      def clipWhenLowerLimitIsLessThanHigher(outputScaledValue, outputRange):
          if (outputScaledValue < outputRange[0]):
              return outputRange[0]
          elif (outputScaledValue > outputRange[1]):
              return outputRange[1]
          else:
              return outputScaledValue
          end
      end

      slope = computeSlope(rawRange, scaledRange)
      intercept = computeIntercept(slope, rawRange, scaledRange)
      scaledValue = slope * value + intercept
      return clipScaledValue(scaledValue, scaledRange)
  end

  def limit(value, range):
      return scale(value, range, range)
  end


  rq_init_comm_if_connected(9, "1")
  rq_init_comm_if_connected(2, "2")
  rq_init_comm_if_connected(3, "3")
  rq_init_comm_if_connected(4, "4")
  rq_print_connected_grippers()
  rq_gripper_communication_thread = run rq_gripper_communication()
  set_closed_norm(97.6470588235294, 1)
  set_open_norm(1.1764705882352942, 1)
  set_closed_mm(0.0, 1)
  set_open_mm(53.0, 1)
  set_closed_norm(100.0, 2)
  set_open_norm(0.0, 2)
  set_closed_mm(0.0, 2)
  set_open_mm(50.0, 2)
  set_closed_norm(100.0, 3)
  set_open_norm(0.0, 3)
  set_closed_mm(0.0, 3)
  set_open_mm(50.0, 3)
  set_closed_norm(100.0, 4)
  set_open_norm(0.0, 4)
  set_closed_mm(0.0, 4)
  set_open_mm(50.0, 4)
  rq_current_limit_enabled = False
  while(not rq_gripper_communication_thread_started):
      sync()
  end
  # end: URCap Installation Node
  # begin: URCap Installation Node
  #   Source: OPC UA, 2.0.2, Rocketfarm AS
  #   Type: OPC UA
  global opcua_daemon = rpc_factory("xmlrpc", "http://127.0.0.1:40409/RPC2")
  def opcua_client_connect(address):
  return opcua_daemon.client_connect(address)
  end
  def opcua_client_get_id(client_name):
  return opcua_daemon.client_get_id(client_name)
  end
  def opcua_client_try_connect(client_id):
  opcua_result = False
  if (opcua_daemon.client_connect(client_id)):
  sleep(0.01)
  opcua_result = opcua_daemon.client_is_connected(client_id)
  opcua_retry = 10
  while ( (not opcua_result) and (opcua_retry > 0) ):
  sleep(0.1)
  opcua_result = opcua_daemon.client_is_connected(client_id)
  opcua_retry = opcua_retry - 1
  end
  end
  return opcua_result
  end
  def opcua_client_disconnect(client_id):
  return opcua_daemon.client_disconnect(client_id)
  end
  def opcua_client_is_connected(client_id):
  return opcua_daemon.client_is_connected(client_id)
  end
  def opcua_client_read_byid(client_id, namespace_id, variable_id):
  return opcua_daemon.client_read_variable_by_id(client_id, namespace_id, variable_id)
  end
  def opcua_client_read_byname(client_id, namespace_id, variable_name):
  return opcua_daemon.client_read_variable_by_name(client_id, namespace_id, variable_name)
  end
  def opcua_client_write_byid(client_id, namespace_id, variable_id, variable_value):
  return opcua_daemon.client_write_variable_by_id(client_id, namespace_id, variable_id, variable_value)
  end
  def opcua_client_write_byname(client_id, namespace_id, variable_name, variable_value):
  return opcua_daemon.client_write_variable_by_name(client_id, namespace_id, variable_name, variable_value)
  end
  def opcua_client_last_error(client_id):
  return opcua_daemon.client_get_last_error(client_id)
  end
  def opcua_server_read_byname(variable_name):
  return opcua_daemon.server_read_variable_by_name(variable_name)
  end
  def opcua_server_write_byname(variable_name, variable_value):
  return opcua_daemon.server_write_variable_by_name(variable_name, variable_value)
  end
  def opcua_server_last_error():
  return opcua_daemon.server_get_last_error()
  end
  def opcua_error_to_string(errorCode):
  return opcua_daemon.error_code_to_string(errorCode)
  end
  # end: URCap Installation Node
  global AMR_Position=struct(position_identifier=0, x1=0, x2=0, y1=0, y2=0, theta1=0, theta2=0)
  global CAM_Pose=p[0,0,0,0,0,0]
  global CAM_Relation=""
  global CMD_Abort=  False
  global CMD_Clear=  False
  global CMD_Reset=  False
  global CMD_Start=  False
  global CMD_Suspend=  False
  global CMD_Unhold=  False
  global CMD_Unsuspend=  False
  global CNT_Rack_Output=0
  global FNC_Freedrive=  False
  global PRC_TubCounter=0
  global STP=0
  global easyPickCount=0
  global easyPickCount_4=0
  global easyPickCount_6=0
  global easyPickNoObj=0
  global easyPickNoObj_4=0
  global easyPickNoObj_6=0
  global easyPickParts=0
  global easyPickParts_4=0
  global easyPickParts_6=0
  global Container_mid_1_p=p[-.379239199143, -.127191311915, .299999999998, .000000000046, -.000000000021, -1.247199999994]
  global Container_mid_1_q=[-2.477408934449926, -1.2969853503591224, -1.875639182904262, -1.539621866126728, 1.5731943360401213, -2.8009955944022717]
  global Container_capt_p=p[-.525590029047, .407247642794, .411588185841, -.000000000107, .000000000065, -2.896148821900]
  global Container_capt_q=[-3.5968351615224767, -2.0050156108707204, -0.8176271154495112, -1.8895759482008394, 1.5730967555598792, -2.2743681102957645]
  global Waypoint_51_p=p[-.335468094724, -.217855817953, .299999999998, .000000000047, -.000000000014, -.994837065669]
  global Waypoint_51_q=[-2.2250460001249586, -1.2969853503591224, -1.875639182904262, -1.539621866126728, 1.573194336040121, -2.800995594402271]
  global Waypoint_65_p=p[-.380578560601, .136229906820, .300065486591, .002668209125, -.001950299791, -1.918285884015]
  global Waypoint_65_q=[-3.1484482924090784, -1.309784547691681, -1.8656262159347534, -1.5396564540318032, 1.5732260942459106, -2.8009706179248255]
  global Waypoint_86_p=p[-.610891912545, .328076512140, .154928874949, -.144389774448, 2.158207980619, -2.101916875088]
  global Waypoint_86_q=[-3.0298424402820032, -2.1616608105101527, -1.770405888557434, -1.8800016842284144, -0.04927570024599248, -0.4936583677874964]
  global Waypoint_16_p=p[-.530358413935, .418971000515, -.109643658887, -.463059997969, 2.087871459122, -2.058033430549]
  global Waypoint_16_q=[-3.2300904432879847, -2.6409207783141078, -1.877760410308838, -1.6937691173949183, -0.43063193956484014, 0.029483795166015625]
  global Waypoint_87_p=p[-.459488806274, .188986755628, .171097942578, -.348072585494, -2.059579317749, 2.019661285019]
  global Waypoint_87_q=[-2.790591303502218, -2.152559896508688, -1.6884642839431763, -2.469414850274557, 0.6884214878082275, 0.021232735365629196]
  global Waypoint_89_p=p[-.261886355761, -.111669623901, .131097242659, -1.173634433322, -1.227274747052, 1.193766216763]
  global Waypoint_89_q=[-2.672995464666928, -2.175407175402028, -1.7617490112425536, -2.338843663300132, 2.030865036219133, 0.036428578240585985]
  global Waypoint_90_p=p[-.269165142951, -.108082457315, .026677271969, -1.173634433324, -1.227274747052, 1.193766216762]
  global Waypoint_90_q=[-2.6853380119023815, -2.380020912479904, -1.7522585114443245, -2.1436252765786143, 2.018787725064888, 0.03659425986402358]
  global Waypoint_88_p=p[-.617446503519, .392270291627, .170489198955, -.224010410006, -2.066036920971, 2.088909130040]
  global Waypoint_88_q=[-3.1488035953258766, -2.4221038789008897, -1.1666724558911366, -2.618578428321003, 0.2380794033913185, -0.04528854192806264]
  global Waypoint_94_p=p[-.452978066378, .173533334300, .109390198136, -.002578830757, -2.196586508502, 2.177068753404]
  global Waypoint_94_q=[-2.6674557574892073, -2.1212895090252317, -1.967198705482553, -2.208419381150989, 0.5117897724834828, 0.04481344519449531]
  global Waypoint_93_p=p[-.596468537907, .142788156334, .105779109453, -.673355127215, 1.831389627653, -1.853156743314]
  global Waypoint_93_q=[-2.6921545586066635, -2.073966887503291, -2.065600898968258, -2.154852607781155, -0.22224352987151796, 0.042304121657345886]
  global Waypoint_95_p=p[-.605386387448, -.069660570533, .218481828695, .000812734400, .006677866481, -1.958478278110]
  global Waypoint_95_q=[-2.8029143834677903, -1.8400819882842256, -1.544169955118452, -1.327224466208456, 1.5676652012497132, -2.4155226342256775]
  global Waypoint_13_p=p[-.479450777041, .284140798427, .125270103493, -.276792173670, 2.098433187455, -2.121256516887]
  global Waypoint_13_q=[-2.8915050665484827, -1.9549266300597132, -2.2318272590637207, -1.6654960117735804, 0.020810842514038086, -0.4019392172442835]
  global Waypoint_70_p=p[-.472820924464, .292439826304, .207418370234, -.259787347864, -2.053484648504, 2.070709755662]
  global Waypoint_70_q=[-2.969927421603815, -2.07168115810532, -1.6835546062719366, -2.4953958198513964, 0.4489790927922641, -0.005578998612037367]
  global Waypoint_2_p=p[-.312961047461, -.152991312519, .223609826854, -.745314530454, -1.713873240489, 1.673341715282]
  global Waypoint_2_q=[-2.3560472170459192, -2.183784624139303, -1.4583134651184082, -2.6435262165465296, 1.6522362232208252, 0.043451953679323196]
  global Waypoint_3_p=p[-.113749865836, -.390110151572, .317307487562, -.519383711706, -.839884211339, 1.756868173041]
  global Waypoint_3_q=[-1.8909733931170862, -1.720626016656393, -1.5115610361099243, -2.1240560017027796, 2.1809096336364746, 0.7227501273155212]
  global Waypoint_15_p=p[.029144035010, -.436802470887, .327885032028, -.521560953301, -.623641814548, 1.862659450154]
  global Waypoint_15_q=[-1.564817253743307, -1.556895188321807, -1.6826975345611572, -1.6944714985289515, 2.2362685203552246, 1.117417335510254]
  global Waypoint_14_p=p[.068712235638, -.569419545175, .285215357659, -.679242949116, -.712065334485, 1.394044574094]
  global Waypoint_14_q=[-1.5731792953485346, -1.8029235103747094, -1.6781008808776736, -1.2218450646111982, 2.4719572998240125, 1.6394218026856375]
  global Waypoint_4_p=p[-.047220457210, -.557624911767, .136370962514, -.679242949107, -.712065334475, 1.394044574096]
  global Waypoint_4_q=[-1.7740079055958748, -2.0023561428872334, -1.7577251142892676, -1.18903287716154, 2.4487287370345143, 1.322902469273079]
  global Waypoint_25_p=p[.065436479647, -.569388431626, .287820755049, -.679242949185, -.712065334557, 1.394044574070]
  global Waypoint_25_q=[-1.5789263550890595, -1.8020194754825436, -1.6702557537748035, -1.237882536889547, 2.471995808083492, 1.6301087487321393]
  global Waypoint_39_p=p[.137772150180, -.577759956854, .299999999946, .000000000217, -.000000000207, -1.594351842625]
  global Waypoint_39_q=[-1.108978697428574, -1.776486680444405, -1.413737665315093, -1.5218908901738937, 1.5733062372356947, -1.0863866394180182]
  global Waypoint_41_p=p[.074222967010, -.565641640647, .234620140366, -.516884386806, .529223682286, -1.529619060506]
  global Waypoint_41_q=[-0.9596722604286052, -1.8767069964135548, -1.4892746174057256, -1.7813862040292285, 1.0520698599867686, -0.8199687448260349]
  global Waypoint_40_p=p[.039987741677, -.564832865048, .191055405868, -.767560686167, .343136533060, -2.241315728308]
  global Waypoint_40_q=[-1.0070649180116558, -1.8745927522477324, -1.6139175023195245, -1.6337474788493545, 1.032708081143138, -0.11587278312988403]
  global Waypoint_42_p=p[.041363380882, -.564865360786, .192805844739, .278500165520, .624117100927, .762272396553]
  global Waypoint_42_q=[-1.0050718976263102, -1.8744386685524779, -1.609151451954446, -1.6399653140247947, 1.0334006002355505, -3.254032861659603]
  global Waypoint_43_p=p[.041363380886, -.564865360780, .192805844755, .854271020883, .226833028600, 2.453002871494]
  global Waypoint_43_q=[-1.0050567614299233, -1.874341297657562, -1.6092945416026048, -1.6397580431809713, 1.0333661149462194, -5.0371728933995605]
  global Waypoint_44_p=p[.040882892233, -.564854254876, .192193763716, .110913882012, .659173708659, .275719738520]
  global Waypoint_44_q=[-1.0057704811530535, -1.8745207681598055, -1.6107765025572558, -1.637858394640876, 1.033164860873599, -2.7487836132940755]
  global Waypoint_45_p=p[.042647731639, -.564895808997, .194439423694, -.451694728506, .563172064821, -1.343350300184]
  global Waypoint_45_q=[-1.0032860829914387, -1.8741561795270565, -1.6048483308761785, -1.6453689714776623, 1.0342050634514657, -1.06078829880322]
  global Waypoint_46_p=p[.099944144487, -.566244126804, .267342790130, -.451694834765, .563172023386, -1.343350532536]
  global Waypoint_46_q=[-0.9257438092434924, -1.889970530402497, -1.3828165217629076, -1.8916791100652528, 1.0664350961373816, -0.9805910833329659]
  global Waypoint_47_p=p[.099944144444, -.566244126727, .267342790273, -.101742139519, .058679218003, -1.457888523314]
  global Waypoint_47_q=[-1.1112623176383014, -1.729989471869196, -1.5530029871033957, -1.4442770617454777, 1.4670579052775654, -1.2224020460061675]
  global Waypoint_48_p=p[-.136182767566, -.647487115908, .294247768372, -.101742139549, .058679218020, -1.457888523312]
  global Waypoint_48_q=[-1.532196177857717, -1.9115932455375173, -1.2651848069729779, -1.5055651746702665, 1.4703193777418382, -1.646379689188814]
  global Waypoint_49_p=p[-.159024328559, -.641021381179, .047691706070, -.000000000033, -.000000000027, -1.457897102937]
  global Waypoint_49_q=[-1.6098490079965062, -2.1164987141784586, -1.6156631902166785, -0.9800092198841526, 1.573231151532669, -1.722204302767242]
  global Waypoint_50_p=p[-.159024328558, -.641021381151, .291114489351, -.000000000033, -.000000000027, -1.457897102937]
  global Waypoint_50_q=[-1.609190265995684, -1.9426985888940234, -1.2189094859258596, -1.55056435122874, 1.5734384912955113, -1.7235116759964022]
  def Sub_Vision_V18():
    $ 650 "Sub_Vision_V18" "noBreak"
    $ 651 "PreSettings"
    $ 652 "CAM_LM_Detected≔ False "
    global CAM_LM_Detected=  False
    $ 653 "CAM_Captures≔0"
    global CAM_Captures=0
    $ 654 "CAM_Pose≔p[0,0,0,0,0,0]"
    global CAM_Pose=p[0,0,0,0,0,0]
    $ 655 "CAM_LM_Refinmnt≔ False "
    global CAM_LM_Refinmnt=  False
    $ 656 "CAM_LM_Refined≔ False "
    global CAM_LM_Refined=  False
    $ 657 "CAM_LM_Deviatn≔p[0,0,0,0,0,0]"
    global CAM_LM_Deviatn=p[0,0,0,0,0,0]
    $ 658 "CAM_LM_ID≔0"
    global CAM_LM_ID=0
    $ 659 "CAM_Done≔ False "
    global CAM_Done=  False
    $ 660 "CAM_CNT_Obj≔0"
    global CAM_CNT_Obj=0
    $ 661 "CAM_Result = []"
    CAM_Result = []
    $ 662 "OBJ_Detected≔ False "
    global OBJ_Detected=  False
    $ 663 "FRM_Reference≔p[0,0,0,0,0,0]"
    global FRM_Reference=p[0,0,0,0,0,0]
    $ 664 "'=========='"
    # '=========='
    $ 665 "Switch Action"
    switch_1 = Action
    $ 666 "Case 13"
    if (13 == switch_1):
    elif (15 == switch_1):
      $ 784 "Case 15"
    elif (131 == switch_1):
      $ 830 "Case 131"
      $ 831 "Read (SensoPart)"
      $ 832 "Action_Info≔'search for landmark'"
      global Action_Info="search for landmark"
      $ 833 "CAM_LM≔CAM_LMs[4]"
      global CAM_LM=CAM_LMs[4]
      $ 834 "CAM_Relation≔CAM_LM.capture_relation"
      global CAM_Relation=CAM_LM.capture_relation
      $ 835 "go to capture pose"
      $ 838 "If ITM_ID≟1 and JIG≟7"
      if (ITM_ID == 1  and  JIG == 7):
        $ 839 "PSE_T≔uLM_Cap_SSRack"
        global PSE_T=uLM_Cap_SSRack
      else:
        $ 840 "ElseIf ITM_ID≟5 and JIG≟7"
        if (ITM_ID == 5  and  JIG == 7):
          $ 841 "PSE_T≔FRM_Cap_SSRack"
          global PSE_T=FRM_Cap_SSRack
        else:
          $ 842 "ElseIf ITM_ID≟13 and JIG≟7"
          if (ITM_ID == 13  and  JIG == 7):
            $ 843 "PSE_T≔FRM_pick_rack_const"
            global PSE_T=p[-0.5568395192387274,0.34423986364170267,0.44698620470146266,-1.0069110132199915E-6,3.378712467497258E-5,-8.002029546773325E-6]
          else:
            $ 844 "ElseIf ITM_ID≟1 and JIG≟15"
            if (ITM_ID == 1 and JIG == 15):
              $ 845 "MoveJ"
              $ 846 "Container_mid_1" "breakAfter"
              movej(get_inverse_kin(Container_mid_1_p, qnear=Container_mid_1_q), a=1.3962634015954636, v=1.0471975511965976, r=0.05)
              $ 847 "Container_capt" "breakAfter"
              movej(get_inverse_kin(Container_capt_p, qnear=Container_capt_q), a=1.3962634015954636, v=1.0471975511965976)
              $ 848 "PSE_T≔FRM_Container_S_const"
              global PSE_T=p[-0.510412665574981,0.40064363362973565,0.41159789496794374,-1.1370875604168537E-5,-3.643547521609506E-6,-2.896122366208473]
            else:
              $ 849 "ElseIf ITM_ID≟1 and JIG≟16"
              if (ITM_ID == 1  and  JIG == 16):
                $ 850 "MoveJ"
                $ 851 "Waypoint_51" "breakAfter"
                movej(get_inverse_kin(Waypoint_51_p, qnear=Waypoint_51_q), a=1.3962634015954636, v=1.0471975511965976, r=0.05)
                $ 854 "PSE_T≔FRM_Container_S_const"
                global PSE_T=p[-0.510412665574981,0.40064363362973565,0.41159789496794374,-1.1370875604168537E-5,-3.643547521609506E-6,-2.896122366208473]
              else:
                $ 855 "ElseIf ITM_ID≟1 and JIG≟17"
                if (ITM_ID == 1  and  JIG == 17):
                  $ 856 "MoveJ"
                  $ 857 "Waypoint_51" "breakAfter"
                  movej(get_inverse_kin(Waypoint_51_p, qnear=Waypoint_51_q), a=1.3962634015954636, v=1.0471975511965976, r=0.05)
                  $ 860 "PSE_T≔FRM_Container_S_const"
                  global PSE_T=p[-0.510412665574981,0.40064363362973565,0.41159789496794374,-1.1370875604168537E-5,-3.643547521609506E-6,-2.896122366208473]
                else:
                  $ 861 "ElseIf ITM_ID≟1 and JIG≟18"
                  if (ITM_ID == 1  and  JIG == 18):
                    $ 864 "MoveJ"
                    $ 865 "Waypoint_51" "breakAfter"
                    movej(get_inverse_kin(Waypoint_51_p, qnear=Waypoint_51_q), a=1.3962634015954636, v=1.0471975511965976, r=0.05)
                    $ 866 "Waypoint_65" "breakAfter"
                    movej(get_inverse_kin(Waypoint_65_p, qnear=Waypoint_65_q), a=1.3962634015954636, v=1.0471975511965976)
                    $ 867 "PSE_T≔FRM_Container_S_const"
                    global PSE_T=p[-0.510412665574981,0.40064363362973565,0.41159789496794374,-1.1370875604168537E-5,-3.643547521609506E-6,-2.896122366208473]
                  else:
                    $ 868 "ElseIf ITM_ID≟1 and JIG≟19"
                    if (ITM_ID == 1  and  JIG == 19):
                      $ 871 "MoveJ"
                      $ 872 "Waypoint_51" "breakAfter"
                      movej(get_inverse_kin(Waypoint_51_p, qnear=Waypoint_51_q), a=1.3962634015954636, v=1.0471975511965976, r=0.05)
                      $ 874 "PSE_T≔aq_rack1_const"
                      global PSE_T=p[-0.6171199234912242,0.18274496130308399,0.4990241423073791,7.867082192074154E-6,-3.513408957609815E-5,-2.5093516385827686]
                    end
                  end
                end
              end
            end
          end
        end
      end
      $ 875 "do_transition(PSE_T, keep_rxry=False)"
      do_transition(PSE_T, keep_rxry=False)
      $ 876 "Set"
      set_tcp(p[0.0,0.0,0.161,3.1415,0.0,0.0])
      $ 877 "MoveJ"
      $ 878 "PSE_T" "breakAfter"
      movej(PSE_T, a=1.3962634015954636, v=1.7453292519943295)
      $ 879 "CAM_Pose≔get_actual_tcp_pose()"
      global CAM_Pose= get_actual_tcp_pose ()
      $ 880 "Loop  not CAM_Done and  not ERROR.FLAG and  not CMD_Stop"
      while (  not  CAM_Done  and    not  ERROR.FLAG  and    not  CMD_Stop):
        $ 881 "adjust capture pose"
        $ 882 "If CAM_LM_Detected and CAM_LM_Refinmnt"
        if (CAM_LM_Detected  and  CAM_LM_Refinmnt):
          $ 883 "PSE_T≔p[0,0,0.300,0,0,0]"
          global PSE_T=p[0,0,0.300,0,0,0]
          $ 884 "CAM_Pose≔PSE_T"
          global CAM_Pose=PSE_T
          $ 885 "If  not is_reachable(FRM_Reference,[PSE_T])"
          if (  not  is_reachable(FRM_Reference,[PSE_T])):
            $ 886 "Error"
            $ 887 "set_error(ERROR_POSE_NOT_REACHABLE)"
            set_error(ERROR_POSE_NOT_REACHABLE)
          end
          $ 888 "If  not ERROR.FLAG"
          if (  not  ERROR.FLAG):
            $ 889 "MoveJ"
            $ 890 "PSE_T" "breakAfter"
            set_tcp(p[0.0,0.0,0.161,0.0,0.0,0.0])
            movej(pose_trans(FRM_Reference, PSE_T), a=0.8726646259971648, v=1.3962634015954636)
            $ 891 "CAM_LM_Refined≔ True "
            global CAM_LM_Refined=  True
          end
        else:
          $ 892 "ElseIf  not CAM_LM_Detected and CAM_Captures>0"
          if (  not  CAM_LM_Detected  and  CAM_Captures>0):
            $ 893 "MoveL"
            $ 894 "If FRM_Reference≟p[0,0,0,0,0,0]"
            if (FRM_Reference == p[0,0,0,0,0,0]):
              $ 895 "PSE_T≔get_random_pose(pose_ref=CAM_Pose, mode='cubic', range_max=[0.150,0.150,0.015])"
              global PSE_T=get_random_pose(pose_ref=CAM_Pose, mode="cubic", range_max=[0.150,0.150,0.015])
            else:
              $ 900 "Else" "noBreak"
              $ 901 "PSE_T≔get_random_pose(pose_ref=CAM_Pose, mode='rotation', range_max=[10,10,0])"
              global PSE_T=get_random_pose(pose_ref=CAM_Pose, mode="rotation", range_max=[10,10,0])
              $ 902 "CAM_LM_Refined≔ True "
              global CAM_LM_Refined=  True
            end
            $ 903 "If get_inverse_kin_has_solution(pose_trans(FRM_Reference, PSE_T))"
            if (get_inverse_kin_has_solution( pose_trans (FRM_Reference, PSE_T))):
              $ 904 "Comment"
              # Comment
              $ 905 "PSE_T" "breakAfter"
              set_tcp(p[0.0,0.0,0.161,3.1415,0.0,0.0])
              movel(pose_trans(FRM_Reference, PSE_T), a=0.03, v=0.05)
            else:
              $ 906 "Else" "noBreak"
              $ 907 "'If random pose is out of reach, set the initial cam pose'"
              # 'If random pose is out of reach, set the initial cam pose'
              $ 908 "PSE_T≔CAM_Pose"
              global PSE_T=CAM_Pose
            end
          end
        end
        $ 909 "Wait: 2.0"
        sleep(2.0)
        $ 910 "trigger"
        $ 911 "If ITM_ID≟1 and JIG≟7"
        if (ITM_ID == 1  and  JIG == 7):
          # begin: URCap Program Node
          #   Source: SensoPart VISOR Robotic, 2.0.0, SensoPart Industriesensorik GmbH
          #   Type: VISOR Trigger
          $ 912 "# 1 VISOR Trigger"
          visor_changeJob(1, "Landmark_INVITE_2", 6000)
          visor_trigger(1, 6000, "arm")
          # end: URCap Program Node
        else:
          $ 913 "ElseIf ITM_ID≟5 and JIG≟7"
          if (ITM_ID == 5  and  JIG == 7):
            # begin: URCap Program Node
            #   Source: SensoPart VISOR Robotic, 2.0.0, SensoPart Industriesensorik GmbH
            #   Type: VISOR Trigger
            $ 914 "# 1 VISOR Trigger"
            visor_changeJob(1, "Landmark_INVITE_2", 6000)
            visor_trigger(1, 6000, "arm")
            # end: URCap Program Node
          else:
            $ 915 "ElseIf ITM_ID≟13 and JIG≟7"
            if (ITM_ID == 13  and  JIG == 7):
              # begin: URCap Program Node
              #   Source: SensoPart VISOR Robotic, 2.0.0, SensoPart Industriesensorik GmbH
              #   Type: VISOR Trigger
              $ 916 "# 1 VISOR Trigger"
              visor_changeJob(1, "Landmark_INVITE_2", 6000)
              visor_trigger(1, 6000, "arm")
              # end: URCap Program Node
            else:
              $ 917 "ElseIf ITM_ID≟1 and JIG≟15"
              if (ITM_ID == 1 and JIG == 15):
                # begin: URCap Program Node
                #   Source: SensoPart VISOR Robotic, 2.0.0, SensoPart Industriesensorik GmbH
                #   Type: VISOR Trigger
                $ 918 "# 1 VISOR Trigger"
                visor_changeJob(1, "PowderA", 6000)
                visor_trigger(1, 6000, "arm")
                # end: URCap Program Node
              else:
                $ 919 "ElseIf ITM_ID≟1 and JIG≟16"
                if (ITM_ID == 1 and JIG == 16):
                  # begin: URCap Program Node
                  #   Source: SensoPart VISOR Robotic, 2.0.0, SensoPart Industriesensorik GmbH
                  #   Type: VISOR Trigger
                  $ 920 "# 1 VISOR Trigger"
                  visor_changeJob(1, "Weigh_target", 6000)
                  visor_trigger(1, 6000, "arm")
                  # end: URCap Program Node
                else:
                  $ 921 "ElseIf ITM_ID≟1 and JIG≟17"
                  if (ITM_ID == 1 and JIG == 17):
                    # begin: URCap Program Node
                    #   Source: SensoPart VISOR Robotic, 2.0.0, SensoPart Industriesensorik GmbH
                    #   Type: VISOR Trigger
                    $ 922 "# 1 VISOR Trigger"
                    visor_changeJob(1, "Weigh_dispense", 6000)
                    visor_trigger(1, 6000, "arm")
                    # end: URCap Program Node
                  else:
                    $ 923 "ElseIf ITM_ID≟1 and JIG≟18"
                    if (ITM_ID == 1 and JIG == 18):
                      # begin: URCap Program Node
                      #   Source: SensoPart VISOR Robotic, 2.0.0, SensoPart Industriesensorik GmbH
                      #   Type: VISOR Trigger
                      $ 924 "# 1 VISOR Trigger"
                      visor_changeJob(1, "pick_rack", 6000)
                      visor_trigger(1, 6000, "arm")
                      # end: URCap Program Node
                    else:
                      $ 926 "ElseIf ITM_ID≟1 and JIG≟19"
                      if (ITM_ID == 1 and JIG == 19):
                        # begin: URCap Program Node
                        #   Source: SensoPart VISOR Robotic, 2.0.0, SensoPart Industriesensorik GmbH
                        #   Type: VISOR Trigger
                        $ 927 "# 1 VISOR Trigger"
                        visor_changeJob(1, "place_rack", 6000)
                        visor_trigger(1, 6000, "arm")
                        # end: URCap Program Node
                      end
                    end
                  end
                end
              end
            end
          end
        end
        $ 932 "TM_3D≔visor_partsFound(1)"
        global TM_3D= visor_partsFound (1)
        $ 933 "If TM_3D>0"
        if (TM_3D>0):
          $ 934 "CAM_LM_Detected≔ True "
          global CAM_LM_Detected=  True
          $ 935 "CAM_Captures≔0"
          global CAM_Captures=0
        else:
          $ 936 "Else" "noBreak"
          $ 937 "CAM_LM_Detected≔ False "
          global CAM_LM_Detected=  False
          $ 938 "CAM_Captures≔CAM_Captures+1"
          global CAM_Captures=CAM_Captures+1
        end
        $ 943 "result"
        $ 944 "If CAM_LM_Detected"
        if (CAM_LM_Detected):
          $ 945 "If (CAM_LM_Refinmnt and CAM_LM_Refined) or  not CAM_LM_Refinmnt"
          if ((CAM_LM_Refinmnt  and  CAM_LM_Refined)  or    not  CAM_LM_Refinmnt):
            $ 1003 "If ITM_ID≟1 and JIG≟7"
            if (ITM_ID == 1  and  JIG == 7):
              $ 1004 "CAM_LM_SSRack≔visor_getPose3d(1, 0)"
              global CAM_LM_SSRack= visor_getPose3d (1, 0)
            else:
              $ 1005 "ElseIf ITM_ID≟5 and JIG≟7"
              if (ITM_ID == 5  and  JIG == 7):
                $ 1006 "CAM_LM_SSRack≔visor_getPose3d(1, 0)"
                global CAM_LM_SSRack= visor_getPose3d (1, 0)
              else:
                $ 1007 "ElseIf ITM_ID≟13 and JIG≟7"
                if (ITM_ID == 13  and  JIG == 7):
                  $ 1008 "CAM_LM_Bott≔visor_getPose3d(1, 0)"
                  global CAM_LM_Bott= visor_getPose3d (1, 0)
                else:
                  $ 1009 "ElseIf ITM_ID≟1 and JIG≟15"
                  if (ITM_ID == 1 and JIG == 15):
                    $ 1010 "CAM_LM_Cont_S≔visor_getPose3d(1, 0)"
                    global CAM_LM_Cont_S= visor_getPose3d (1, 0)
                    $ 1011 "cont_img_pose≔get_actual_tcp_pose()"
                    global cont_img_pose= get_actual_tcp_pose ()
                  else:
                    $ 1012 "ElseIf ITM_ID≟1 and JIG≟16"
                    if (ITM_ID == 1 and JIG == 16):
                      $ 1013 "CAM_cont≔visor_getPose3d(1, 0)"
                      global CAM_cont= visor_getPose3d (1, 0)
                      $ 1014 "cont_img_pose≔get_actual_tcp_pose()"
                      global cont_img_pose= get_actual_tcp_pose ()
                    else:
                      $ 1015 "ElseIf ITM_ID≟1 and JIG≟17"
                      if (ITM_ID == 1 and JIG == 17):
                        $ 1016 "pose_rack_aq1≔visor_getPose3d(1, 0)"
                        global pose_rack_aq1= visor_getPose3d (1, 0)
                        $ 1017 "cont_img_pose≔get_actual_tcp_pose()"
                        global cont_img_pose= get_actual_tcp_pose ()
                      else:
                        $ 1018 "ElseIf ITM_ID≟1 and JIG≟18"
                        if (ITM_ID == 1 and JIG == 18):
                          $ 1019 "pose_rack_aq1≔visor_getPose3d(1, 0)"
                          global pose_rack_aq1= visor_getPose3d (1, 0)
                          $ 1020 "FRM_Container_S≔get_actual_tcp_pose()"
                          global FRM_Container_S= get_actual_tcp_pose ()
                        else:
                          $ 1021 "ElseIf ITM_ID≟1 and JIG≟19"
                          if (ITM_ID == 1 and JIG == 19):
                            $ 1022 "pose_rack_aq1≔visor_getPose3d(1, 0)"
                            global pose_rack_aq1= visor_getPose3d (1, 0)
                            $ 1023 "aq_rack1≔get_actual_tcp_pose()"
                            global aq_rack1= get_actual_tcp_pose ()
                          end
                        end
                      end
                    end
                  end
                end
              end
            end
            $ 1024 "CAM_Done≔ True "
            global CAM_Done=  True
          end
        else:
          $ 1025 "ElseIf  not CAM_LM_Detected and CAM_Captures<CAM_PRM_Retries"
          if (  not  CAM_LM_Detected  and  CAM_Captures<CAM_PRM_Retries):
            $ 1026 "CAM_LM_Refined≔ False "
            global CAM_LM_Refined=  False
          else:
            $ 1027 "ElseIf CAM_Captures≥CAM_PRM_Retries"
            if (CAM_Captures >= CAM_PRM_Retries):
              $ 1028 "CAM_Done≔ True "
              global CAM_Done=  True
              $ 1029 "Error"
              $ 1030 "set_error(ERROR_NO_LANDMARK)"
              set_error(ERROR_NO_LANDMARK)
            end
          end
        end
      end
    elif (151 == switch_1):
      $ 1031 "Case 151"
      $ 1032 "Detect (SensoPart)"
      $ 1033 "go to capture pose"
      $ 1034 "FRM_Reference≔FRM_Cap_SSRack"
      global FRM_Reference=FRM_Cap_SSRack
      $ 1035 "PSE_T≔p[0,0,-0.00,0,0,0]"
      global PSE_T=p[0,0,-0.00,0,0,0]
      $ 1036 "do_transition(pose_trans(FRM_Reference, PSE_T), keep_rxry=False)"
      do_transition( pose_trans (FRM_Reference, PSE_T), keep_rxry=False)
      $ 1037 "JNT_Q≔get_actual_joint_positions()"
      global JNT_Q= get_actual_joint_positions ()
      $ 1038 "JNT_Q≔[JNT_Q[0], JNT_Q[1], JNT_Q[2], JNT_Q[3], JNT_Q[4], 0]"
      global JNT_Q=[JNT_Q[0], JNT_Q[1], JNT_Q[2], JNT_Q[3], JNT_Q[4], 0]
      $ 1039 "Set"
      set_tcp(p[0.0,0.0,0.161,3.1415,0.0,0.0])
      $ 1040 "movej(get_inverse_kin(pose_trans(FRM_Reference, PSE_T), qnear=JNT_Q))"
      movej(get_inverse_kin( pose_trans (FRM_Reference, PSE_T), qnear=JNT_Q))
      $ 1041 "CAM_Pose≔pose_trans(pose_inv(FRM_Reference), get_actual_tcp_pose())"
      global CAM_Pose= pose_trans ( pose_inv (FRM_Reference),  get_actual_tcp_pose ())
      $ 1042 "Loop  not CAM_Done and  not ERROR.FLAG and  not CMD_Stop"
      while (  not  CAM_Done  and    not  ERROR.FLAG  and    not  CMD_Stop):
        $ 1043 "If  not OBJ_Detected and CAM_Captures>0"
        if (  not  OBJ_Detected  and  CAM_Captures>0):
          $ 1044 "MoveL"
          $ 1045 "If FRM_Reference≟p[0,0,0,0,0,0]"
          if (FRM_Reference == p[0,0,0,0,0,0]):
            $ 1047 "PSE_T≔get_random_pose(pose_ref=CAM_Pose, mode='rotation', range_max=[15,15,0])"
            global PSE_T=get_random_pose(pose_ref=CAM_Pose, mode="rotation", range_max=[15,15,0])
          else:
            $ 1048 "Else" "noBreak"
            $ 1049 "PSE_T≔get_random_pose(pose_ref=CAM_Pose, mode='rotation', range_max=[10,10,0])"
            global PSE_T=get_random_pose(pose_ref=CAM_Pose, mode="rotation", range_max=[10,10,0])
          end
          $ 1050 "If get_inverse_kin_has_solution(pose_trans(FRM_Reference, PSE_T))"
          if (get_inverse_kin_has_solution( pose_trans (FRM_Reference, PSE_T))):
            $ 1051 "PSE_T" "breakAfter"
            set_tcp(p[0.0,0.0,0.161,3.1415,0.0,0.0])
            movel(pose_trans(FRM_Reference, PSE_T), a=0.03, v=0.05)
          else:
            $ 1052 "Else" "noBreak"
            $ 1053 "'If random pose is out of reach, set the initial cam pose'"
            # 'If random pose is out of reach, set the initial cam pose'
            $ 1054 "PSE_T≔CAM_Pose"
            global PSE_T=CAM_Pose
            $ 1055 "PSE_T" "breakAfter"
            set_tcp(p[0.0,0.0,0.161,3.1415,0.0,0.0])
            movel(pose_trans(FRM_Reference, PSE_T), a=0.03, v=0.05)
          end
        end
        $ 1056 "Wait: 0.5"
        sleep(0.5)
        $ 1057 "Set"
        set_tcp(p[0.0,0.0,0.161,3.1415,0.0,0.0])
        # begin: URCap Program Node
        #   Source: SensoPart VISOR Robotic, 2.0.0, SensoPart Industriesensorik GmbH
        #   Type: VISOR Trigger
        $ 1058 "# 1 VISOR Trigger"
        visor_changeJob(1, "Object Detection Single", 6000)
        visor_trigger(1, 6000, "arm")
        # end: URCap Program Node
        $ 1059 "If visor_isResponseOk(1)"
        if ( visor_isResponseOk (1)):
          $ 1060 "CAM_CNT_Obj≔visor_partsFound(1)"
          global CAM_CNT_Obj= visor_partsFound (1)
          $ 1061 "CAM_OBJ_Pose≔visor_getPose3d(1, 0)"
          global CAM_OBJ_Pose= visor_getPose3d (1, 0)
          $ 1062 "If CAM_CNT_Obj>0"
          if (CAM_CNT_Obj>0):
            $ 1063 "CAM_OBJ_Color≔visor_getAdditionalData(1, 0)"
            global CAM_OBJ_Color= visor_getAdditionalData (1, 0)
            $ 1064 "CAM_DetectScore≔to_num(visor_getAdditionalData(1, 1))/1000"
            global CAM_DetectScore=to_num( visor_getAdditionalData (1, 1))/1000
            $ 1065 "OBJ_Detected≔ True "
            global OBJ_Detected=  True
          end
        else:
          $ 1066 "Else" "noBreak"
          $ 1067 "CAM_Captures≔CAM_Captures+1"
          global CAM_Captures=CAM_Captures+1
        end
        $ 1068 "If OBJ_Detected"
        if (OBJ_Detected):
          $ 1069 "Get object data"
          $ 1070 "PRC_CntDetect≔0"
          global PRC_CntDetect=0
          $ 1071 "Loop PRC_CntDetect<CAM_CNT_Obj"
          while (PRC_CntDetect<CAM_CNT_Obj):
            $ 1072 "get object and jig number"
            $ 1073 "If ITM_ID≟1 and JIG≟7"
            if (ITM_ID == 1  and  JIG == 7):
              $ 1074 "FRM_Reference≔FRM_Cap_SSRack"
              global FRM_Reference=FRM_Cap_SSRack
            else:
              $ 1075 "ElseIf ITM_ID≟5 and JIG≟7"
              if (ITM_ID == 5  and  JIG == 7):
                $ 1076 "FRM_Reference≔uLM_Cap_SSRack"
                global FRM_Reference=uLM_Cap_SSRack
              end
            end
            $ 1079 "PSE_T≔pose_trans(pose_inv(FRM_Reference), CAM_OBJ_Pose)"
            global PSE_T= pose_trans ( pose_inv (FRM_Reference), CAM_OBJ_Pose)
            $ 1080 "CAM_Result.append(get_pattern_counter(PSE_T, 'X', pattern=[10, 5], patternsize=[0.181, 0.081]))"
            CAM_Result.append(get_pattern_counter(PSE_T, "X", pattern=[10, 5], patternsize=[0.181, 0.081]))
            $ 1081 "PRC_CntDetect≔PRC_CntDetect+1"
            global PRC_CntDetect=PRC_CntDetect+1
          end
          $ 1082 "CAM_Done≔ True "
          global CAM_Done=  True
        else:
          $ 1083 "ElseIf CAM_Captures≥CAM_PRM_Retries"
          if (CAM_Captures >= CAM_PRM_Retries):
            $ 1084 "CAM_Done≔ True "
            global CAM_Done=  True
          else:
            $ 1085 "Else" "noBreak"
            $ 1086 "CAM_Captures≔CAM_Captures+1"
            global CAM_Captures=CAM_Captures+1
          end
        end
      end
    end
    $ 1087 "'=========='"
    # '=========='
    $ 1088 "PostSettings"
    $ 1089 "FRM_Reference≔p[0,0,0,0,0,0]"
    global FRM_Reference=p[0,0,0,0,0,0]
    $ 1090 "Set"
    set_tcp(p[0.0,0.0,0.161,3.1415,0.0,0.0])
    $ 1091 "CAM_Pose≔p[0,0,0,0,0,0]"
    global CAM_Pose=p[0,0,0,0,0,0]
    $ 1092 "Action≔0"
    global Action=0
    $ 1093 "Action_Info≔''"
    global Action_Info=""
  end
  def Sub_AMR_MiR_V3():
    $ 1094 "Sub_AMR_MiR_V3" "noBreak"
    $ 1095 "PreSettings"
    $ 1096 "AMR_TargetList≔[1,2,3,4,5,21,22,23,24,31,32,33,34,35,36,37,38,41]"
    global AMR_TargetList=[1,2,3,4,5,21,22,23,24,31,32,33,34,35,36,37,38,41]
    $ 1097 "AMR_Done≔ False "
    global AMR_Done=  False
    $ 1098 "AMR_PosActual≔T2O_Current_Pos"
    global AMR_PosActual=modbus_get_signal_status("T2O_Current_Pos")
    $ 1099 "AMR_Attemps≔T2O_Nav_Attemps"
    global AMR_Attemps=modbus_get_signal_status("T2O_Nav_Attemps")
    $ 1100 "AMR_Battery≔MiR_Battery_Lvl"
    global AMR_Battery=modbus_get_signal_status("MiR_Battery_Lvl")
    $ 1101 "AMR_Charging≔(T2O_Charging≟1)"
    global AMR_Charging=(modbus_get_signal_status("T2O_Charging") == 1)
    $ 1102 "AMR_Position≔struct(position_identifier=T2O_Current_Pos, x1=MiR_Position_X1, x2=MiR_Position_X2, y1=MiR_Position_Y1, y2=MiR_Position_Y2, theta1=MiR_Theta_1, theta2=MiR_Theta_2) "
    global AMR_Position=struct(position_identifier=modbus_get_signal_status("T2O_Current_Pos"), x1=modbus_get_signal_status("MiR_Position_X1"), x2=modbus_get_signal_status("MiR_Position_X2"), y1=modbus_get_signal_status("MiR_Position_Y1"), y2=modbus_get_signal_status("MiR_Position_Y2"), theta1=modbus_get_signal_status("MiR_Theta_1"), theta2=modbus_get_signal_status("MiR_Theta_2"))
    $ 1103 "If MiR_Mode≠7"
    if (modbus_get_signal_status("MiR_Mode") != 7):
      $ 1104 "Error"
      $ 1105 "set_error(ERROR_AMR_WRONG_MODE)"
      set_error(ERROR_AMR_WRONG_MODE)
      $ 1106 "AMR_Done≔ True "
      global AMR_Done=  True
    end
    $ 1107 "'=========='"
    # '=========='
    $ 1108 "Switch STATE"
    switch_1 = STATE
    $ 1109 "Case 1"
    if (1 == switch_1):
      $ 1110 "stopping"
      $ 1111 "If T2O_Done≟1 and O2T_Acknowledge≟0"
      if (modbus_get_signal_status("T2O_Done") == 1  and  modbus_get_signal_status("O2T_Acknowledge") == 0):
        $ 1112 "Set O2T_Acknowledge=1"
        modbus_set_output_register("O2T_Acknowledge", 1)
      end
      $ 1113 "Set MiR_CMD_Stop=On"
      modbus_set_output_signal("MiR_CMD_Stop", True)
      $ 1114 "AMR_Position.position_identifier = 0"
      AMR_Position.position_identifier = 0
      $ 1115 "AMR_Done≔ True "
      global AMR_Done=  True
    elif (2 == switch_1):
      $ 1116 "Case 2"
      $ 1117 "stopped"
      $ 1118 "If MiR_State≠3 and MiR_State≠5"
      if (modbus_get_signal_status("MiR_State") != 3  and  modbus_get_signal_status("MiR_State") != 5):
        $ 1119 "Set MiR_CMD_Stop=Off"
        modbus_set_output_signal("MiR_CMD_Stop", False)
      end
    elif (3 == switch_1):
      $ 1120 "Case 3"
      $ 1121 "resetting"
      $ 1122 "Set O2T_Mis_Main=Off"
      modbus_set_output_signal("O2T_Mis_Main", False)
      $ 1123 "Set O2T_Mis_Charge=Off"
      modbus_set_output_signal("O2T_Mis_Charge", False)
      $ 1124 "If MiR_Mis_Queue>0"
      if (modbus_get_signal_status("MiR_Mis_Queue")>0):
        $ 1125 "Set MiR_CMD_Clear_Q=On"
        modbus_set_output_signal("MiR_CMD_Clear_Q", True)
        $ 1126 "Wait MiR_Mis_Queue≟0"
        while (not(modbus_get_signal_status("MiR_Mis_Queue") == 0)):
          sync()
        end
        $ 1127 "Set MiR_CMD_Clear_Q=Off"
        modbus_set_output_signal("MiR_CMD_Clear_Q", False)
      end
      $ 1128 "If MiR_Error_ID≠0"
      if (modbus_get_signal_status("MiR_Error_ID") != 0):
        $ 1129 "Set MiR_CMD_Clear_E=On"
        modbus_set_output_signal("MiR_CMD_Clear_E", True)
        $ 1130 "Wait MiR_Error_ID≟0"
        while (not(modbus_get_signal_status("MiR_Error_ID") == 0)):
          sync()
        end
        $ 1131 "Set MiR_CMD_Clear_E=Off"
        modbus_set_output_signal("MiR_CMD_Clear_E", False)
      end
      $ 1132 "Set O2T_Action=0"
      modbus_set_output_register("O2T_Action", 0)
      $ 1133 "Set O2T_Acknowledge=0"
      modbus_set_output_register("O2T_Acknowledge", 0)
      $ 1134 "Set O2T_Target_Pos=0"
      modbus_set_output_register("O2T_Target_Pos", 0)
      $ 1135 "Set O2T_Footprint=0"
      modbus_set_output_register("O2T_Footprint", 0)
      $ 1136 "Set O2T_ProtectOff=0"
      modbus_set_output_register("O2T_ProtectOff", 0)
      $ 1137 "Set O2T_Dock=0"
      modbus_set_output_register("O2T_Dock", 0)
      $ 1138 "AMR_Attemps≔0"
      global AMR_Attemps=0
      $ 1139 "AMR_PosTarget≔0"
      global AMR_PosTarget=0
      $ 1140 "AMR_Step≔0"
      global AMR_Step=0
      $ 1141 "AMR_AtTarget≔ False "
      global AMR_AtTarget=  False
      $ 1142 "If MiR_State≟4 or MiR_State≟3 or MiR_State≟10"
      if (modbus_get_signal_status("MiR_State") == 4  or  modbus_get_signal_status("MiR_State") == 3  or  modbus_get_signal_status("MiR_State") == 10):
        $ 1143 "AMR_Done≔ True "
        global AMR_Done=  True
      end
    elif (5 == switch_1):
      $ 1144 "Case 5"
      $ 1145 "starting"
      $ 1146 "If MiR_State≟4"
      if (modbus_get_signal_status("MiR_State") == 4):
        $ 1147 "Set MiR_CMD_Start=On"
        modbus_set_output_signal("MiR_CMD_Start", True)
        $ 1148 "Wait MiR_State≠4"
        while (not(modbus_get_signal_status("MiR_State") != 4)):
          sync()
        end
        $ 1149 "Set MiR_CMD_Start=Off"
        modbus_set_output_signal("MiR_CMD_Start", False)
        $ 1150 "AMR_Done≔ True "
        global AMR_Done=  True
      else:
        $ 1151 "ElseIf MiR_State≟10"
        if (modbus_get_signal_status("MiR_State") == 10):
          $ 1152 "'MiR in protective stop. Wait'"
          # 'MiR in protective stop. Wait'
          $ 1153 "AMR_Done≔ True "
          global AMR_Done=  True
        else:
          $ 1154 "ElseIf MiR_State≟3"
          if (modbus_get_signal_status("MiR_State") == 3):
            $ 1155 "AMR_Done≔ True "
            global AMR_Done=  True
          end
        end
      end
    elif (6 == switch_1):
      $ 1156 "Case 6"
      $ 1157 "execute"
      $ 1158 "AMR_AtTarget≔(AMR_PosActual≟AMR_PosTarget)"
      global AMR_AtTarget=(AMR_PosActual == AMR_PosTarget)
      $ 1159 "Switch AMR_Step"
      switch_2 = AMR_Step
      $ 1160 "Case 0"
      if (0 == switch_2):
        $ 1161 "If  not AMR_AtTarget"
        if (  not  AMR_AtTarget):
          $ 1162 "AMR_Step≔1"
          global AMR_Step=1
        else:
          $ 1163 "Else" "noBreak"
          $ 1164 "AMR_Done≔ True "
          global AMR_Done=  True
        end
      elif (1 == switch_2):
        $ 1165 "Case 1"
        $ 1166 "general Settings"
        $ 1167 "Set O2T_Acknowledge=0"
        modbus_set_output_register("O2T_Acknowledge", 0)
        $ 1168 "check for error"
        $ 1169 "If OBJ_Picked and MiR_State≟10"
        if (OBJ_Picked  and  modbus_get_signal_status("MiR_State") == 10):
          $ 1170 "Error"
          $ 1171 "set_error(ERROR_ROBOT_ARM_NOT_IN_HOME_POSE)"
          set_error(ERROR_ROBOT_ARM_NOT_IN_HOME_POSE)
          $ 1172 "Action≔0"
          global Action=0
        else:
          $ 1173 "ElseIf  not found_in_list(AMR_PosTarget, AMR_TargetList)"
          if (  not  found_in_list(AMR_PosTarget, AMR_TargetList)):
            $ 1174 "Error"
            $ 1175 "set_error(ERROR_UNKNOWN_POSE)"
            set_error(ERROR_UNKNOWN_POSE)
            $ 1176 "Action≔0"
            global Action=0
          end
        end
        $ 1177 "If MiR_State≟3"
        if (modbus_get_signal_status("MiR_State") == 3):
          $ 1178 "Set MiR_CMD_Start=Off"
          modbus_set_output_signal("MiR_CMD_Start", False)
          $ 1179 "Switch Action"
          switch_3 = Action
          $ 1180 "Case 51"
          if (51 == switch_3):
            $ 1181 "Charge"
            $ 1182 "'trigger the charging mission'"
            # 'trigger the charging mission'
            $ 1183 "'target pos is predefined'"
            # 'target pos is predefined'
            $ 1184 "Set O2T_Footprint=0"
            modbus_set_output_register("O2T_Footprint", 0)
            $ 1185 "Set O2T_Action=1"
            modbus_set_output_register("O2T_Action", 1)
            $ 1186 "If MiR_Mis_Queue≟0"
            if (modbus_get_signal_status("MiR_Mis_Queue") == 0):
              $ 1187 "Set O2T_Mis_Charge=On"
              modbus_set_output_signal("O2T_Mis_Charge", True)
              $ 1188 "Wait MiR_Mis_Queue≥1"
              while (not(modbus_get_signal_status("MiR_Mis_Queue") >= 1)):
                sync()
              end
              $ 1189 "Set O2T_Mis_Charge=Off"
              modbus_set_output_signal("O2T_Mis_Charge", False)
            end
          elif (52 == switch_3):
            $ 1190 "Case 52"
            $ 1191 "Navigate"
            $ 1192 "'trigger the standard missoin'"
            # 'trigger the standard missoin'
            $ 1193 "Set O2T_Footprint=AMR_FootprintID"
            modbus_set_output_register("O2T_Footprint", AMR_FootprintID)
            $ 1194 "Set O2T_Target_Pos=AMR_PosTarget"
            modbus_set_output_register("O2T_Target_Pos", AMR_PosTarget)
            $ 1195 "Set O2T_Action=2"
            modbus_set_output_register("O2T_Action", 2)
            $ 1196 "If MiR_Mis_Queue≟0"
            if (modbus_get_signal_status("MiR_Mis_Queue") == 0):
              $ 1197 "Set O2T_Mis_Main=On"
              modbus_set_output_signal("O2T_Mis_Main", True)
              $ 1198 "Wait MiR_Mis_Queue≥1"
              while (not(modbus_get_signal_status("MiR_Mis_Queue") >= 1)):
                sync()
              end
              $ 1199 "Set O2T_Mis_Main=Off"
              modbus_set_output_signal("O2T_Mis_Main", False)
            end
          end
        else:
          $ 1200 "ElseIf MiR_State≟4"
          if (modbus_get_signal_status("MiR_State") == 4):
            $ 1201 "Set MiR_CMD_Start=On"
            modbus_set_output_signal("MiR_CMD_Start", True)
          else:
            $ 1202 "ElseIf MiR_State≟5"
            if (modbus_get_signal_status("MiR_State") == 5):
              $ 1203 "AMR_Step≔2"
              global AMR_Step=2
            else:
              $ 1204 "ElseIf MiR_State≟10"
              if (modbus_get_signal_status("MiR_State") == 10):
                $ 1205 "'AMR still in safeguard stop'"
                # 'AMR still in safeguard stop'
              end
            end
          end
        end
      elif (2 == switch_2):
        $ 1206 "Case 2"
        $ 1207 "acknowledge handshake"
        $ 1208 "If T2O_Done≟1 and O2T_Acknowledge≟0"
        if (modbus_get_signal_status("T2O_Done") == 1  and  modbus_get_signal_status("O2T_Acknowledge") == 0):
          $ 1209 "Set O2T_Acknowledge=1"
          modbus_set_output_register("O2T_Acknowledge", 1)
        else:
          $ 1210 "ElseIf T2O_Done≟0 and O2T_Acknowledge≟1"
          if (modbus_get_signal_status("T2O_Done") == 0  and  modbus_get_signal_status("O2T_Acknowledge") == 1):
            $ 1211 "Set O2T_Acknowledge=0"
            modbus_set_output_register("O2T_Acknowledge", 0)
            $ 1212 "AMR_AtTarget≔(AMR_PosActual≟AMR_PosTarget)"
            global AMR_AtTarget=(AMR_PosActual == AMR_PosTarget)
            $ 1213 "AMR_Done≔ True "
            global AMR_Done=  True
          end
        end
      end
      $ 1214 "translate errors"
      $ 1215 "If AMR_Done"
      if (AMR_Done):
        $ 1216 "Switch T2O_Error_ID"
        switch_2 = modbus_get_signal_status("T2O_Error_ID")
        $ 1217 "Case 2003"
        if (2003 == switch_2):
          $ 1218 "error"
          $ 1219 "set_error(ERROR_NOT_DOCKED)"
          set_error(ERROR_NOT_DOCKED)
        elif (2007 == switch_2):
          $ 1220 "Case 2007"
          $ 1221 "error"
          $ 1222 "set_error(ERROR_NOT_REACHABLE_TARGET)"
          set_error(ERROR_NOT_REACHABLE_TARGET)
        elif (2008 == switch_2):
          $ 1223 "Case 2008"
          $ 1224 "error"
          $ 1225 "set_error(ERROR_CHARGING_NOT_STARTED)"
          set_error(ERROR_CHARGING_NOT_STARTED)
        end
      end
    elif (7 == switch_1):
      $ 1226 "Case 7"
      $ 1227 "completing"
      $ 1228 "If MiR_Mis_Queue>0"
      if (modbus_get_signal_status("MiR_Mis_Queue")>0):
        $ 1229 "Set MiR_CMD_Abort=On"
        modbus_set_output_signal("MiR_CMD_Abort", True)
        $ 1230 "Wait MiR_Mis_Queue≟0"
        while (not(modbus_get_signal_status("MiR_Mis_Queue") == 0)):
          sync()
        end
        $ 1231 "Set MiR_CMD_Abort=Off"
        modbus_set_output_signal("MiR_CMD_Abort", False)
      end
      $ 1232 "If MiR_State≟3 or MiR_State≟10"
      if (modbus_get_signal_status("MiR_State") == 3  or  modbus_get_signal_status("MiR_State") == 10):
        $ 1233 "AMR_Done≔ True "
        global AMR_Done=  True
      end
    elif (9 == switch_1):
      $ 1234 "Case 9"
      $ 1235 "holding"
      $ 1236 "Set MiR_CMD_Abort=On"
      modbus_set_output_signal("MiR_CMD_Abort", True)
      $ 1237 "If MiR_State≟3 or MiR_State≟10"
      if (modbus_get_signal_status("MiR_State") == 3  or  modbus_get_signal_status("MiR_State") == 10):
        $ 1238 "Set MiR_CMD_Abort=Off"
        modbus_set_output_signal("MiR_CMD_Abort", False)
        $ 1239 "AMR_Done≔ True "
        global AMR_Done=  True
      end
    elif (11 == switch_1):
      $ 1240 "Case 11"
      $ 1241 "unholding"
      $ 1242 "Set MiR_CMD_Start=On"
      modbus_set_output_signal("MiR_CMD_Start", True)
      $ 1243 "If MiR_State≠4"
      if (modbus_get_signal_status("MiR_State") != 4):
        $ 1244 "Set MiR_CMD_Start=Off"
        modbus_set_output_signal("MiR_CMD_Start", False)
        $ 1245 "AMR_Step≔0"
        global AMR_Step=0
        $ 1246 "AMR_Done≔ True "
        global AMR_Done=  True
      end
    elif (12 == switch_1):
      $ 1247 "Case 12"
      $ 1248 "suspending"
      $ 1249 "'none'"
      # 'none'
    elif (14 == switch_1):
      $ 1250 "Case 14"
      $ 1251 "unsuspending"
      $ 1252 "'none'"
      # 'none'
    elif (15 == switch_1):
      $ 1253 "Case 15"
      $ 1254 "aborting"
      $ 1255 "Set MiR_CMD_Abort=On"
      modbus_set_output_signal("MiR_CMD_Abort", True)
      $ 1256 "Wait MiR_State≟3"
      while (not(modbus_get_signal_status("MiR_State") == 3)):
        sync()
      end
      $ 1257 "Set MiR_CMD_Abort=Off"
      modbus_set_output_signal("MiR_CMD_Abort", False)
    elif (17 == switch_1):
      $ 1258 "Case 17"
      $ 1259 "clearing"
      $ 1260 "If MiR_Error_ID≠0"
      if (modbus_get_signal_status("MiR_Error_ID") != 0):
        $ 1261 "Set MiR_CMD_Clear_E=On"
        modbus_set_output_signal("MiR_CMD_Clear_E", True)
        $ 1262 "Wait MiR_Error_ID≟0"
        while (not(modbus_get_signal_status("MiR_Error_ID") == 0)):
          sync()
        end
        $ 1263 "Set MiR_CMD_Clear_E=Off"
        modbus_set_output_signal("MiR_CMD_Clear_E", False)
      end
      $ 1264 "If MiR_Error_ID≟0"
      if (modbus_get_signal_status("MiR_Error_ID") == 0):
        $ 1265 "AMR_Done≔ True "
        global AMR_Done=  True
      end
    end
    $ 1266 "'=========='"
    # '=========='
    $ 1267 "PostSettings"
    $ 1268 "AMR_Position≔struct(position_identifier=T2O_Current_Pos, x1=MiR_Position_X1, x2=MiR_Position_X2, y1=MiR_Position_Y1, y2=MiR_Position_Y2, theta1=MiR_Theta_1, theta2=MiR_Theta_2) "
    global AMR_Position=struct(position_identifier=modbus_get_signal_status("T2O_Current_Pos"), x1=modbus_get_signal_status("MiR_Position_X1"), x2=modbus_get_signal_status("MiR_Position_X2"), y1=modbus_get_signal_status("MiR_Position_Y1"), y2=modbus_get_signal_status("MiR_Position_Y2"), theta1=modbus_get_signal_status("MiR_Theta_1"), theta2=modbus_get_signal_status("MiR_Theta_2"))
  end
  def Sub_Action_V4():
    $ 1269 "Sub_Action_V4" "noBreak"
    $ 1270 "PreSettings"
    $ 1271 "init poses"
    $ 1272 "PSE_A≔p[0,0,0,0,0,0]"
    global PSE_A=p[0,0,0,0,0,0]
    $ 1273 "PSE_A_H≔p[0,0,0,0,0,0]"
    global PSE_A_H=p[0,0,0,0,0,0]
    $ 1274 "PSE_T≔p[0,0,0,0,0,0]"
    global PSE_T=p[0,0,0,0,0,0]
    $ 1275 "PSE_T_H≔p[0,0,0,0,0,0]"
    global PSE_T_H=p[0,0,0,0,0,0]
    $ 1276 "PSE_G≔p[0,0,0,0,0,0]"
    global PSE_G=p[0,0,0,0,0,0]
    $ 1277 "PSE_G_H≔p[0,0,0,0,0,0]"
    global PSE_G_H=p[0,0,0,0,0,0]
    $ 1278 "PSE_R≔p[0,0,0,0,0,0]"
    global PSE_R=p[0,0,0,0,0,0]
    $ 1279 "PSE_R_H≔p[0,0,0,0,0,0]"
    global PSE_R_H=p[0,0,0,0,0,0]
    $ 1280 "JNT_Q≔[0,0,0,0,0,0]"
    global JNT_Q=[0,0,0,0,0,0]
    $ 1281 "JNT_S≔[0,0,0,0,0,0]"
    global JNT_S=[0,0,0,0,0,0]
    $ 1282 "Gripping parameters"
    $ 1283 "OBJ = find_object_by_type(OBJs, OBJ_Type)"
    OBJ = find_object_by_type(OBJs, OBJ_Type)
    $ 1284 "GRP_Open_Pos≔OBJ.dimension.diameter * 1000 + 6"
    global GRP_Open_Pos=OBJ.dimension.diameter * 1000 + 6
    $ 1285 "GRP_Offset≔OBJ.gripper_offset"
    global GRP_Offset=OBJ.gripper_offset
    $ 1286 "rq_set_force_norm(50)"
     rq_set_force_norm (50)
    $ 1287 "rq_set_speed_norm(50)"
     rq_set_speed_norm (50)
    $ 1288 "Switch ITM_ID"
    switch_1 = ITM_ID
    $ 1289 "Case 1"
    if (1 == switch_1):
      $ 1290 "uML"
      $ 1291 "JIG2 = find_object_by_type(JIGs, JIG)"
      JIG2 = find_object_by_type(JIGs, JIG)
      $ 1292 "JIG_Offset≔JIG2.jig_offset"
      global JIG_Offset=JIG2.jig_offset
      $ 1293 "Switch JIG"
      switch_2 = JIG
      $ 1294 "Case 1"
      if (1 == switch_2):
        $ 1295 "3FG"
        $ 1296 "define poses"
        $ 1297 "FRM_Reference≔ULM_3FG"
        global FRM_Reference=ULM_3FG
        $ 1298 "JNT_Q≔JNT_HOME"
        global JNT_Q=JNT_HOME
        $ 1299 "PSE_T≔pose_trans(GRP_Offset, JIG_Offset)"
        global PSE_T= pose_trans (GRP_Offset, JIG_Offset)
        $ 1300 "PSE_A≔pose_trans(PSE_T, p[0,0,0.100,0,0,0])"
        global PSE_A= pose_trans (PSE_T, p[0,0,0.100,0,0,0])
        $ 1301 "PSE_R≔pose_add(PSE_T, p[0,0,0.100,0,0,0])"
        global PSE_R= pose_add (PSE_T, p[0,0,0.100,0,0,0])
      elif (2 == switch_2):
        $ 1302 "Case 2"
        $ 1303 "Input"
        $ 1304 "'CHANGE THE REFERENCE TO THE FRAME TO MOVE IN'"
        # 'CHANGE THE REFERENCE TO THE FRAME TO MOVE IN'
        $ 1305 "define poses"
        $ 1306 "FRM_Reference≔ULM_Input"
        global FRM_Reference=ULM_Input
        $ 1307 "PSE_T≔pose_trans(pose_trans(get_pattern_pos_rectangle(OBJ_Nbr, 'X', [10,5], patternsize=[0.181,0.081]), GRP_Offset), JIG_Offset)"
        global PSE_T= pose_trans ( pose_trans (get_pattern_pos_rectangle(OBJ_Nbr, "X", [10,5], patternsize=[0.181,0.081]), GRP_Offset), JIG_Offset)
        $ 1308 "If Action≟1"
        if (Action == 1):
          $ 1309 "PSE_R≔pose_add(PSE_T, p[0,0,0.200,0,0,0])"
          global PSE_R= pose_add (PSE_T, p[0,0,0.200,0,0,0])
          $ 1310 "PSE_A≔pose_add(PSE_T, p[0,0,0.100,0,0,0])"
          global PSE_A= pose_add (PSE_T, p[0,0,0.100,0,0,0])
        else:
          $ 1311 "ElseIf Action≟2"
          if (Action == 2):
            $ 1312 "PSE_R≔pose_add(PSE_T, p[0,0,0.100,0,0,0])"
            global PSE_R= pose_add (PSE_T, p[0,0,0.100,0,0,0])
            $ 1313 "PSE_A≔pose_add(PSE_T, p[0,0,0.200,0,0,0])"
            global PSE_A= pose_add (PSE_T, p[0,0,0.200,0,0,0])
          end
        end
      elif (3 == switch_2):
        $ 1314 "Case 3"
        $ 1315 "Output"
        $ 1316 "'CHANGE THE REFERENCE TO THE FRAME TO MOVE IN'"
        # 'CHANGE THE REFERENCE TO THE FRAME TO MOVE IN'
        $ 1317 "define poses"
        $ 1318 "FRM_Reference≔ULM_Output"
        global FRM_Reference=ULM_Output
        $ 1319 "PSE_T≔pose_trans(pose_trans(get_pattern_pos_rectangle(OBJ_Nbr, 'X', [10,5], patternsize=[0.181,0.081]), GRP_Offset), JIG_Offset)"
        global PSE_T= pose_trans ( pose_trans (get_pattern_pos_rectangle(OBJ_Nbr, "X", [10,5], patternsize=[0.181,0.081]), GRP_Offset), JIG_Offset)
        $ 1321 "If Action≟1"
        if (Action == 1):
          $ 1322 "PSE_R≔pose_add(PSE_T, p[0,0,0.200,0,0,0])"
          global PSE_R= pose_add (PSE_T, p[0,0,0.200,0,0,0])
          $ 1323 "PSE_A≔pose_add(PSE_T, p[0,0,0.100,0,0,0])"
          global PSE_A= pose_add (PSE_T, p[0,0,0.100,0,0,0])
        else:
          $ 1324 "ElseIf Action≟2"
          if (Action == 2):
            $ 1325 "PSE_R≔pose_add(PSE_T, p[0,0,0.100,0,0,0])"
            global PSE_R= pose_add (PSE_T, p[0,0,0.100,0,0,0])
            $ 1326 "PSE_A≔pose_add(PSE_T, p[0,0,0.200,0,0,0])"
            global PSE_A= pose_add (PSE_T, p[0,0,0.200,0,0,0])
          end
        end
      elif (4 == switch_2):
        $ 1327 "Case 4"
        $ 1328 "jig centrifuge racks"
        $ 1329 "define poses"
        $ 1330 "FRM_Reference≔ULM_Cent_Racks"
        global FRM_Reference=ULM_Cent_Racks
        $ 1331 "PSE_T≔get_pattern_pos_rectangle(JIG_Slot, 'X', [4,1], patternsize=[0.291,0])"
        global PSE_T=get_pattern_pos_rectangle(JIG_Slot, "X", [4,1], patternsize=[0.291,0])
        $ 1332 "If OBJ_Nbr≠0"
        if (OBJ_Nbr != 0):
          $ 1333 "PSE_T≔pose_trans(pose_trans(PSE_T, get_pattern_pos_rectangle(OBJ_Nbr, 'X', [3,3], patternsize=[0.060,0.060])),p[-0.030, -0.030,0,0,0,3.927])"
          global PSE_T= pose_trans ( pose_trans (PSE_T, get_pattern_pos_rectangle(OBJ_Nbr, "X", [3,3], patternsize=[0.060,0.060])),p[-0.030, -0.030,0,0,0,3.927])
        end
        $ 1334 "PSE_T≔pose_trans(PSE_T, GRP_Offset)"
        global PSE_T= pose_trans (PSE_T, GRP_Offset)
        $ 1335 "If Action≟1"
        if (Action == 1):
          $ 1336 "PSE_R≔pose_add(PSE_T, p[0,0,0.200,0,0,0])"
          global PSE_R= pose_add (PSE_T, p[0,0,0.200,0,0,0])
          $ 1337 "PSE_A≔pose_add(PSE_T, p[0,0,0.100,0,0,0])"
          global PSE_A= pose_add (PSE_T, p[0,0,0.100,0,0,0])
        else:
          $ 1338 "ElseIf Action≟2"
          if (Action == 2):
            $ 1339 "PSE_R≔pose_add(PSE_T, p[0,0,0.100,0,0,0])"
            global PSE_R= pose_add (PSE_T, p[0,0,0.100,0,0,0])
            $ 1340 "PSE_A≔pose_add(PSE_T, p[0,0,0.200,0,0,0])"
            global PSE_A= pose_add (PSE_T, p[0,0,0.200,0,0,0])
          end
        end
      elif (6 == switch_2):
        $ 1341 "Case 6"
        $ 1342 "Caps bin"
        $ 1343 "define poses"
        $ 1344 "'Drop cap'"
        # 'Drop cap'
        $ 1345 "FRM_Reference=ULM_Cap_Bin"
        FRM_Reference=ULM_Cap_Bin
        $ 1346 "PSE_T≔pose_RPY2RotVec(p[0,0,0,0,0,0])"
        global PSE_T=pose_RPY2RotVec(p[0,0,0,0,0,0])
        $ 1347 "PSE_T_H≔pose_add(PSE_T, p[0,0,-0.011,0,0,0])"
        global PSE_T_H= pose_add (PSE_T, p[0,0,-0.011,0,0,0])
        $ 1348 "PSE_A≔pose_trans(PSE_T, p[0,0,0.1,0,0,0])"
        global PSE_A= pose_trans (PSE_T, p[0,0,0.1,0,0,0])
        $ 1349 "PSE_R_H≔pose_add(PSE_T, p[0,0,0.100,0,0,0])"
        global PSE_R_H= pose_add (PSE_T, p[0,0,0.100,0,0,0])
        $ 1350 "PSE_R≔pose_add(PSE_T, p[0,0,0.100,0,0,0])"
        global PSE_R= pose_add (PSE_T, p[0,0,0.100,0,0,0])
      elif (7 == switch_2):
        $ 1351 "Case 7"
        $ 1352 "Sarstedt"
        $ 1353 "'CHANGE THE REFERENCE TO THE FRAME TO MOVE IN'"
        # 'CHANGE THE REFERENCE TO THE FRAME TO MOVE IN'
        $ 1359 "If TASK.ID≟10"
        if (TASK.ID == 10):
          $ 1360 "Frame & Position Params"
          $ 1362 "FRM_Reference = CAM_LM_SSRack"
          FRM_Reference = CAM_LM_SSRack
          $ 1367 "PSE_T≔uLM_SS_PickPlc"
          global PSE_T=uLM_SS_PickPlc
          $ 1368 "PSE_A≔pose_trans(PSE_T, p[0,0,0.1,0,0,0])"
          global PSE_A= pose_trans (PSE_T, p[0,0,0.1,0,0,0])
          $ 1369 "PSE_R≔pose_add(PSE_T, p[0,0,0.1,0,0,0])"
          global PSE_R= pose_add (PSE_T, p[0,0,0.1,0,0,0])
        else:
          $ 1370 "ElseIf TASK.ID≟11"
          if (TASK.ID == 11):
            $ 1371 "FRM_Reference = ULM_SS_Jig"
            FRM_Reference = ULM_SS_Jig
            $ 1372 "PSE_T≔pose_RPY2RotVec(p[0,0,0,0,0,0])"
            global PSE_T=pose_RPY2RotVec(p[0,0,0,0,0,0])
            $ 1373 "PSE_T≔pose_trans(PSE_T, GRP_Offset)"
            global PSE_T=pose_trans(PSE_T, GRP_Offset)
            $ 1374 "PSE_A≔pose_trans(PSE_T, p[0,0,0.1,0,0,0])"
            global PSE_A= pose_trans (PSE_T, p[0,0,0.1,0,0,0])
            $ 1375 "PSE_R≔pose_add(PSE_T, p[0,0,0.2,0,0,0])"
            global PSE_R= pose_add (PSE_T, p[0,0,0.2,0,0,0])
          end
        end
      elif (8 == switch_2):
        $ 1376 "Case 8"
        $ 1377 "NoK"
        $ 1378 "define poses"
        $ 1379 "'NoK'"
        # 'NoK'
        $ 1380 "FRM_Reference=ULM_NoK"
        FRM_Reference=ULM_NoK
        $ 1381 "PSE_T≔pose_RPY2RotVec(p[0,0,0,0,0,0])"
        global PSE_T=pose_RPY2RotVec(p[0,0,0,0,0,0])
        $ 1382 "PSE_A≔pose_trans(PSE_T, p[0,0,0.1,0,0,0])"
        global PSE_A= pose_trans (PSE_T, p[0,0,0.1,0,0,0])
        $ 1383 "PSE_R≔pose_add(PSE_T, p[0,0,0.100,0,0,0])"
        global PSE_R= pose_add (PSE_T, p[0,0,0.100,0,0,0])
      elif (9 == switch_2):
        $ 1384 "Case 9"
        $ 1385 "Pick_bott_jig"
        $ 1386 "define poses"
        $ 1387 "'NoK'"
        # 'NoK'
        $ 1388 "FRM_Reference=ULM_bottle_pick_const"
        FRM_Reference=p[0.08175869478771049,-0.47602162643540935,0.09,0.00141829700319658,-0.0027789445191063835,0.07763675748118615]
        $ 1389 "PSE_T≔pose_RPY2RotVec(p[0,0,0,0,0,0])"
        global PSE_T=pose_RPY2RotVec(p[0,0,0,0,0,0])
        $ 1390 "PSE_A≔pose_trans(PSE_T, p[0,0,0.1,0,0,0])"
        global PSE_A= pose_trans (PSE_T, p[0,0,0.1,0,0,0])
        $ 1391 "PSE_R≔pose_add(PSE_T, p[0,0,0.100,0,0,0])"
        global PSE_R= pose_add (PSE_T, p[0,0,0.100,0,0,0])
      elif (10 == switch_2):
        $ 1392 "Case 10"
        $ 1393 "Place_bott_jig"
        $ 1394 "define poses"
        $ 1395 "'NoK'"
        # 'NoK'
        $ 1396 "FRM_Reference=ULM_bottle_plac_const"
        FRM_Reference=p[-0.09502738395762109,-0.5154087721098056,0.095,0.0014590126708889871,-0.0028280855286173575,0.07763149296298452]
        $ 1397 "PSE_T≔pose_RPY2RotVec(p[0,0,0,0,0,0])"
        global PSE_T=pose_RPY2RotVec(p[0,0,0,0,0,0])
        $ 1398 "PSE_A≔pose_trans(PSE_T, p[0,0,0.1,0,0,0])"
        global PSE_A= pose_trans (PSE_T, p[0,0,0.1,0,0,0])
        $ 1399 "PSE_R≔pose_add(PSE_T, p[0,0,0.100,0,0,0])"
        global PSE_R= pose_add (PSE_T, p[0,0,0.100,0,0,0])
      elif (11 == switch_2):
        $ 1400 "Case 11"
        $ 1401 "Place_bott_jig"
        $ 1402 "define poses"
        $ 1403 "'NoK'"
        # 'NoK'
        $ 1404 "FRM_Reference=shake"
        FRM_Reference=shake
        $ 1405 "PSE_T≔pose_RPY2RotVec(p[0,0,0,0,0,0])"
        global PSE_T=pose_RPY2RotVec(p[0,0,0,0,0,0])
        $ 1406 "PSE_A≔pose_trans(PSE_T, p[0,0,0,0,0,0])"
        global PSE_A= pose_trans (PSE_T, p[0,0,0,0,0,0])
        $ 1407 "PSE_R≔pose_add(PSE_T, p[0,0,0,0,0,0])"
        global PSE_R= pose_add (PSE_T, p[0,0,0,0,0,0])
      elif (12 == switch_2):
        $ 1408 "Case 12"
        $ 1409 "Pick_Vial_jig"
        $ 1410 "define poses"
        $ 1411 "'NoK'"
        # 'NoK'
        $ 1412 "FRM_Reference=shake"
        FRM_Reference=shake
        $ 1413 "PSE_T≔pose_RPY2RotVec(p[0,0,0,0,0,0])"
        global PSE_T=pose_RPY2RotVec(p[0,0,0,0,0,0])
        $ 1414 "PSE_A≔pose_trans(PSE_T, p[0,0,0,0,0,0])"
        global PSE_A= pose_trans (PSE_T, p[0,0,0,0,0,0])
        $ 1415 "PSE_R≔pose_add(PSE_T, p[0,0,0,0,0,0])"
        global PSE_R= pose_add (PSE_T, p[0,0,0,0,0,0])
      end
    elif (2 == switch_1):
      $ 1416 "Case 2"
      $ 1417 "Centrifuge"
      $ 1418 "'CHANGE THE REFERENCE TO THE FRAME TO MOVE IN'"
      # 'CHANGE THE REFERENCE TO THE FRAME TO MOVE IN'
      $ 1419 "define poses"
      $ 1420 "FRM_Reference≔FRM_Centrifuge"
      global FRM_Reference=FRM_Centrifuge
      $ 1421 "PSE_T≔GRP_Offset"
      global PSE_T=GRP_Offset
      $ 1422 "If Action≟8"
      if (Action == 8):
        $ 1423 "PSE_R≔pose_add(PSE_T, p[0,0,0.250,0,0,0])"
        global PSE_R= pose_add (PSE_T, p[0,0,0.250,0,0,0])
        $ 1424 "PSE_A≔pose_add(PSE_T, p[0,0,0.150,0,0,0])"
        global PSE_A= pose_add (PSE_T, p[0,0,0.150,0,0,0])
      else:
        $ 1425 "ElseIf Action≟7"
        if (Action == 7):
          $ 1426 "PSE_R≔pose_add(PSE_T, p[0,0,0.150,0,0,0])"
          global PSE_R= pose_add (PSE_T, p[0,0,0.150,0,0,0])
          $ 1427 "PSE_A≔pose_add(PSE_T, p[0,0,0.250,0,0,0])"
          global PSE_A= pose_add (PSE_T, p[0,0,0.250,0,0,0])
        end
      end
    elif (3 == switch_1):
      $ 1428 "Case 3"
      $ 1429 "Output"
      $ 1430 "'CHANGE THE REFERENCE TO THE FRAME TO MOVE IN'"
      # 'CHANGE THE REFERENCE TO THE FRAME TO MOVE IN'
      $ 1431 "define poses"
      $ 1432 "FRM_Reference≔Base_const"
      global FRM_Reference=p[0.0,0.0,0.0,0.0,0.0,0.0]
      $ 1433 "PSE_T≔p[0,0,0,0,0,0]"
      global PSE_T=p[0,0,0,0,0,0]
      $ 1434 "PSE_A≔pose_add(PSE_T, p[0,0,0.150,0,0,0])"
      global PSE_A= pose_add (PSE_T, p[0,0,0.150,0,0,0])
      $ 1435 "PSE_R≔pose_add(PSE_T, p[0,0,0.100,0,0,0])"
      global PSE_R= pose_add (PSE_T, p[0,0,0.100,0,0,0])
    elif (5 == switch_1):
      $ 1436 "Case 5"
      $ 1437 "Sarstedt Pickup Table"
      $ 1438 "'CHANGE THE REFERENCE TO THE FRAME TO MOVE IN'"
      # 'CHANGE THE REFERENCE TO THE FRAME TO MOVE IN'
      $ 1439 "Switch JIG"
      switch_2 = JIG
      $ 1440 "Case 7"
      if (7 == switch_2):
        $ 1453 "Sarstedt"
        $ 1454 "'CHANGE THE REFERENCE TO THE FRAME TO MOVE IN'"
        # 'CHANGE THE REFERENCE TO THE FRAME TO MOVE IN'
        $ 1460 "If TASK.ID≟10"
        if (TASK.ID == 10):
          $ 1461 "Frame & Position Params"
          $ 1462 "FRM_Reference = CAM_LM_SSRack"
          FRM_Reference = CAM_LM_SSRack
          $ 1463 "PSE_T≔uLM_SS_PickPlc"
          global PSE_T=uLM_SS_PickPlc
          $ 1464 "PSE_A≔pose_trans(PSE_T, p[0,0,0.1,0,0,0])"
          global PSE_A= pose_trans (PSE_T, p[0,0,0.1,0,0,0])
          $ 1465 "PSE_R≔pose_add(PSE_T, p[0,0,0.1,0,0,0])"
          global PSE_R= pose_add (PSE_T, p[0,0,0.1,0,0,0])
        end
      end
    elif (13 == switch_1):
      $ 1472 "Case 13"
      $ 1473 "Sarstedt Pickup Table"
      $ 1474 "'CHANGE THE REFERENCE TO THE FRAME TO MOVE IN'"
      # 'CHANGE THE REFERENCE TO THE FRAME TO MOVE IN'
      $ 1475 "Switch JIG"
      switch_2 = JIG
      $ 1476 "Case 7"
      if (7 == switch_2):
        $ 1489 "Bottle"
        $ 1490 "'CHANGE THE REFERENCE TO THE FRAME TO MOVE IN'"
        # 'CHANGE THE REFERENCE TO THE FRAME TO MOVE IN'
        $ 1496 "If TASK.ID≟43"
        if (TASK.ID == 43):
          $ 1497 "Frame & Position Params"
          $ 1498 "FRM_Reference = CAM_LM_Bott"
          FRM_Reference = CAM_LM_Bott
          $ 1499 "PSE_T≔uLM_SS_PickPlc"
          global PSE_T=uLM_SS_PickPlc
          $ 1500 "PSE_A≔pose_trans(PSE_T, p[0,0,0.1,0,0,0])"
          global PSE_A= pose_trans (PSE_T, p[0,0,0.1,0,0,0])
          $ 1501 "PSE_R≔pose_add(PSE_T, p[0,0,0.1,0,0,0])"
          global PSE_R= pose_add (PSE_T, p[0,0,0.1,0,0,0])
        end
      end
    end
    $ 1508 "Additional check"
    $ 1509 "If  not is_reachable(FRM_Reference,[PSE_A,PSE_A_H,PSE_T,PSE_T_H,PSE_R,PSE_R_H])"
    if (  not  is_reachable(FRM_Reference,[PSE_A,PSE_A_H,PSE_T,PSE_T_H,PSE_R,PSE_R_H])):
      $ 1510 "Error"
      $ 1511 "set_error(ERROR_POSE_NOT_REACHABLE)"
      set_error(ERROR_POSE_NOT_REACHABLE)
      $ 1512 "Action≔0"
      global Action=0
    end
    $ 1513 "'=========='"
    # '=========='
    $ 1514 "Switch Action"
    switch_1 = Action
    $ 1515 "Case 1"
    if (1 == switch_1):
      $ 1516 "Pick"
      $ 1517 "Action_Info≔'pick object'"
      global Action_Info="pick object"
      $ 1518 "do_transition(pose_trans(FRM_Reference, PSE_T), keep_rxry=OBJ_Picked)"
      do_transition( pose_trans (FRM_Reference, PSE_T), keep_rxry=OBJ_Picked)
      $ 1519 "EOAT"
      $ 1520 "If  not OBJ_Picked"
      if (  not  OBJ_Picked):
        $ 1521 "rq_move_and_wait_mm(GRP_Open_Pos)"
         rq_move_and_wait_mm (GRP_Open_Pos)
      end
      $ 1522 "If PSE_A_H≠PSE_Z"
      if (PSE_A_H != PSE_Z):
        $ 1523 "If JNT_Q≠JNT_Z"
        if (JNT_Q != JNT_Z):
          $ 1524 "movej(get_inverse_kin(pose_trans(FRM_Reference, PSE_A_H), qnear=JNT_Q), r=0.050)"
          movej(get_inverse_kin( pose_trans (FRM_Reference, PSE_A_H), qnear=JNT_Q), r=0.050)
        else:
          $ 1525 "Else" "noBreak"
          $ 1526 "movej(pose_trans(FRM_Reference, PSE_A_H), r=0.050)"
          movej( pose_trans (FRM_Reference, PSE_A_H), r=0.050)
        end
      end
      $ 1527 "If PSE_A≠PSE_Z"
      if (PSE_A != PSE_Z):
        $ 1528 "If JNT_Q≠JNT_Z"
        if (JNT_Q != JNT_Z):
          $ 1529 "movej(get_inverse_kin(pose_trans(FRM_Reference, PSE_A), qnear=JNT_Q), r=0.020)"
          movej(get_inverse_kin( pose_trans (FRM_Reference, PSE_A), qnear=JNT_Q), r=0.020)
        else:
          $ 1530 "Else" "noBreak"
          $ 1531 "movej(pose_trans(FRM_Reference, PSE_A), r=0.020)"
          movej( pose_trans (FRM_Reference, PSE_A), r=0.020)
        end
      end
      $ 1532 "MoveL"
      $ 1533 "If PSE_T_H≠PSE_Z"
      if (PSE_T_H != PSE_Z):
        $ 1534 "PSE_T_H" "breakAfter"
        movel(pose_trans(FRM_Reference, PSE_T_H), a=0.5, v=0.4, r=0.01)
      end
      $ 1535 "PSE_T" "breakAfter"
      movel(pose_trans(FRM_Reference, PSE_T), a=0.08, v=0.12)
      $ 1536 "EOAT"
      $ 1537 "rq_set_force_norm(50)"
       rq_set_force_norm (50)
      $ 1538 "rq_close_and_wait()"
       rq_close_and_wait ()
      $ 1539 "OBJ_Picked≔rq_is_object_detected()"
      global OBJ_Picked= rq_is_object_detected ()
      $ 1540 "If  not OBJ_Picked"
      if (  not  OBJ_Picked):
        $ 1541 "set_error(ERROR_NO_OBJECT_TO_PICK)"
        set_error(ERROR_NO_OBJECT_TO_PICK)
      end
      $ 1542 "EXTT"
      $ 1543 "Switch JIG"
      switch_2 = JIG
      $ 1544 "Case 1"
      if (1 == switch_2):
        $ 1545 "3FG"
        $ 1546 "If OBJ_Picked"
        if (OBJ_Picked):
          $ 1547 "Set GRP_3F_Open=On"
          set_standard_digital_out(5, True)
        end
      end
      $ 1548 "If PSE_R_H≠PSE_Z"
      if (PSE_R_H != PSE_Z):
        $ 1549 "PSE_R" "breakAfter"
        movel(pose_trans(FRM_Reference, PSE_R), a=0.5, v=0.4, r=0.01)
        $ 1550 "PSE_R_H" "breakAfter"
        movel(pose_trans(FRM_Reference, PSE_R_H), a=0.5, v=0.4)
      else:
        $ 1551 "Else" "noBreak"
        $ 1552 "PSE_R" "breakAfter"
        movel(pose_trans(FRM_Reference, PSE_R), a=0.5, v=0.4)
      end
    elif (2 == switch_1):
      $ 1553 "Case 2"
    elif (3 == switch_1):
      $ 1595 "Case 3"
    elif (4 == switch_1):
      $ 1598 "Case 4"
    elif (5 == switch_1):
      $ 1601 "Case 5"
      $ 1602 "Pick the deepwell rack"
      # begin: URCap Program Node
      #   Source: SensoPart VISOR Robotic, 2.0.0, SensoPart Industriesensorik GmbH
      #   Type: VISOR Robotic App
      $ 1603 "VISOR Easy Pick"
      def visorFuncEasyPick_863a74():
        # begin: URCap Program Node
        #   Source: SensoPart VISOR Robotic, 2.0.0, SensoPart Industriesensorik GmbH
        #   Type: Easy Pick Setup
        $ 1604 "# 1 Setup" "noBreak"
        local easyPickVisorId = 1
        local easyPickArmMounted = True
        local easyPickSetJob = True
        local easyPickJobName = "pick_rack"
        local easyPickAtImgAcq = False
        local easyPickImgAcqPose = FRM_Container_S
        # end: URCap Program Node
        # begin: URCap Program Node
        #   Source: SensoPart VISOR Robotic, 2.0.0, SensoPart Industriesensorik GmbH
        #   Type: Process
        $ 1605 "Process" "noBreak"
        local easyPickObjTaken = False
        local easyPickTrigger = False
        local easyPickPoseIdx = 0
        local easyPickPose = p[0,0,0,0,0,0]
        def easyPickFuncTrigger(visorId, setJob, jobName, arm):
        if (setJob):
          visor_changeJob(visorId, jobName, 6000)
        end
        if (arm):
          visor_trigger(visorId, 6000, "arm")
        else:
          visor_trigger(visorId, 6000)
        end
        global easyPickParts=visor_partsFound(visorId)
        visor_easyPickUpdate(visorId, "parts", visor_partsFound(visorId))
        return visor_getPose3d(visorId, 0)
      end
      while (not easyPickObjTaken):
        easyPickTrigger = (easyPickCount >= visor_partsFound(easyPickVisorId)) or (easyPickCount > 9) or (not visor_easyPickCheckIdent("a6c257", easyPickVisorId))
        if (easyPickTrigger):
          easyPickCount = 0
        end
        easyPickPoseIdx = easyPickCount
        easyPickPose = visor_getPose3d(easyPickVisorId, easyPickPoseIdx)
        visor_easyPickUpdate(easyPickVisorId, "counter", easyPickPoseIdx)
        # begin: URCap Program Node
        #   Source: SensoPart VISOR Robotic, 2.0.0, SensoPart Industriesensorik GmbH
        #   Type: Image Acquisition Pose
        $ 1606 "Image Acquisition Pose" "noBreak"
        if (easyPickTrigger):
          if (not easyPickAtImgAcq):
            movej(pose_trans(easyPickImgAcqPose,p[0.0000,0.0000,-0.0000,0.0000,0.0000,0.0000]),a=1.3963,v=1.0472,t=0.000000,r=0.000000)
            easyPickAtImgAcq = True
          end
          easyPickPose = easyPickFuncTrigger(easyPickVisorId, easyPickSetJob, easyPickJobName, easyPickArmMounted)
        end
        # end: URCap Program Node
        # begin: URCap Program Node
        #   Source: SensoPart VISOR Robotic, 2.0.0, SensoPart Industriesensorik GmbH
        #   Type: Object Detected
        $ 1607 "Object Detected" "noBreak"
        if (visor_partsFound(easyPickVisorId) > 0):
          $ 1608 "Open Gripper" "noBreak"
          # begin: URCap Program Node
          #   Source: Robotiq_Grippers, 1.8.4.4844, Robotiq Inc.
          #   Type: Gripper
          $ 1609 "Gripper Open (1)" "noBreak"
          if not(gripper_connected[0]):
            popup("Gripper 1 must be connected to run this program.", "No connection", False, True, True)
          end
          if not(rq_is_gripper_activated("1")):
            popup("Gripper 1 is not activated. Go to Installation tab > Gripper to activate it and run the program again.", "Not activated", False, True, True)
          end
          rq_set_pos_spd_for(0, 102, 77, "1")
          rq_wait_pos_spe_for_request(0, 102, 77, "1")
          rq_go_to("1")
          rq_wait("1")
          # end: URCap Program Node
          $ 1610 "MoveJ" "noBreak"
          $ 1611 "Waypoint_86" "noBreak"
          movej(get_inverse_kin(Waypoint_86_p, qnear=Waypoint_86_q), a=0.6981317007977318, v=0.5235987755982988)
          # begin: URCap Program Node
          #   Source: SensoPart VISOR Robotic, 2.0.0, SensoPart Industriesensorik GmbH
          #   Type: Approach Pose
          $ 1612 "Approach Pose" "noBreak"
          movej(pose_trans(easyPickPose,p[0.0000,0.0000,0.0500,0.0000,0.0000,0.0000]),a=0.6981,v=0.5236,t=0.000000,r=0.000000)
          # end: URCap Program Node
          # begin: URCap Program Node
          #   Source: SensoPart VISOR Robotic, 2.0.0, SensoPart Industriesensorik GmbH
          #   Type: Target Pose
          $ 1613 "Target Pose" "noBreak"
          movel(pose_trans(easyPickPose,p[0.0000,0.0000,-0.0000,0.0000,0.0000,0.0000]),a=0.2000,v=0.1200,t=0.000000,r=0.000000)
          # end: URCap Program Node
          $ 1614 "Close Gripper" "noBreak"
          # begin: URCap Program Node
          #   Source: Robotiq_Grippers, 1.8.4.4844, Robotiq Inc.
          #   Type: Gripper
          $ 1615 "Gripper Close (1)" "noBreak"
          if not(gripper_connected[0]):
            popup("Gripper 1 must be connected to run this program.", "No connection", False, True, True)
          end
          if not(rq_is_gripper_activated("1")):
            popup("Gripper 1 is not activated. Go to Installation tab > Gripper to activate it and run the program again.", "Not activated", False, True, True)
          end
          rq_set_pos_spd_for(255, 102, 77, "1")
          rq_wait_pos_spe_for_request(255, 102, 77, "1")
          rq_go_to("1")
          rq_wait("1")
          # end: URCap Program Node
          # begin: URCap Program Node
          #   Source: SensoPart VISOR Robotic, 2.0.0, SensoPart Industriesensorik GmbH
          #   Type: Exit Pose
          $ 1616 "Exit Pose" "noBreak"
          movel(pose_trans(easyPickPose,p[0.0000,0.0000,-0.0000,0.0000,0.0000,0.0000]),a=0.2000,v=0.1200,t=0.000000,r=0.000000)
          # end: URCap Program Node
          easyPickObjTaken = True
        end
        # end: URCap Program Node
        # begin: URCap Program Node
        #   Source: SensoPart VISOR Robotic, 2.0.0, SensoPart Industriesensorik GmbH
        #   Type: No Object Detected
        $ 1617 "No Object Detected" "noBreak"
        if (visor_partsFound(easyPickVisorId) < 1):
          $ 1618 "Popup: No Container detected" "noBreak"
          popup("No Container detected", "Message", False, False, blocking=True)
          else:
        end
        # end: URCap Program Node
      end
      easyPickCount = easyPickCount + 1
      visor_easyPickUpdate(easyPickVisorId, "counter", easyPickCount)
      visor_easyPickSetIdent("a6c257", easyPickVisorId)
      # end: URCap Program Node
    end
    visorFuncEasyPick_863a74()
    # end: URCap Program Node
    $ 1619 "Wait: 2.0"
    sleep(2.0)
    $ 1620 "MoveJ"
    $ 1621 "Waypoint_16" "breakAfter"
    movej(get_inverse_kin(Waypoint_16_p, qnear=Waypoint_16_q), a=0.6981317007977318, v=0.3490658503988659)
    $ 1622 "Waypoint_87" "breakAfter"
    movej(get_inverse_kin(Waypoint_87_p, qnear=Waypoint_87_q), a=0.6981317007977318, v=0.3490658503988659)
    $ 1623 "Waypoint_89" "breakAfter"
    movej(get_inverse_kin(Waypoint_89_p, qnear=Waypoint_89_q), a=0.6981317007977318, v=0.3490658503988659)
    $ 1624 "MoveL"
    $ 1625 "Waypoint_90" "breakAfter"
    movel(Waypoint_90_p, a=0.6, v=0.12)
    # begin: URCap Program Node
    #   Source: Robotiq_Grippers, 1.8.4.4844, Robotiq Inc.
    #   Type: Gripper
    $ 1626 "Gripper Open (1)"
    if not(gripper_connected[0]):
      popup("Gripper 1 must be connected to run this program.", "No connection", False, True, True)
    end
    if not(rq_is_gripper_activated("1")):
      popup("Gripper 1 is not activated. Go to Installation tab > Gripper to activate it and run the program again.", "Not activated", False, True, True)
    end
    rq_set_pos_spd_for(0, 0, 0, "1")
    rq_wait_pos_spe_for_request(0, 0, 0, "1")
    rq_go_to("1")
    rq_wait("1")
    # end: URCap Program Node
    $ 1627 "Waypoint_89" "breakAfter"
    movel(Waypoint_89_p, a=0.6, v=0.12)
  elif (6 == switch_1):
    $ 1628 "Case 6"
    $ 1643 "offset≔p[0, 0.03, 0, 0, 0, 0]"
    global offset=p[0, 0.03, 0, 0, 0, 0]
    $ 1644 "Place the deepwell rack"
    # begin: URCap Program Node
    #   Source: SensoPart VISOR Robotic, 2.0.0, SensoPart Industriesensorik GmbH
    #   Type: VISOR Robotic App
    $ 1645 "VISOR Easy Pick"
    def visorFuncEasyPick_d789e5():
      # begin: URCap Program Node
      #   Source: SensoPart VISOR Robotic, 2.0.0, SensoPart Industriesensorik GmbH
      #   Type: Easy Pick Setup
      $ 1646 "# 1 Setup" "noBreak"
      local easyPickVisorId = 1
      local easyPickArmMounted = True
      local easyPickSetJob = True
      local easyPickJobName = "place_rack"
      local easyPickAtImgAcq = False
      local easyPickImgAcqPose = aq_rack1
      # end: URCap Program Node
      # begin: URCap Program Node
      #   Source: SensoPart VISOR Robotic, 2.0.0, SensoPart Industriesensorik GmbH
      #   Type: Process
      $ 1647 "Process" "noBreak"
      local easyPickObjTaken = False
      local easyPickTrigger = False
      local easyPickPoseIdx = 0
      local easyPickPose = p[0,0,0,0,0,0]
      def easyPickFuncTrigger(visorId, setJob, jobName, arm):
      if (setJob):
        visor_changeJob(visorId, jobName, 6000)
      end
      if (arm):
        visor_trigger(visorId, 6000, "arm")
      else:
        visor_trigger(visorId, 6000)
      end
      global easyPickParts=visor_partsFound(visorId)
      visor_easyPickUpdate(visorId, "parts", visor_partsFound(visorId))
      return visor_getPose3d(visorId, 0)
    end
    while (not easyPickObjTaken):
      easyPickTrigger = (easyPickCount >= visor_partsFound(easyPickVisorId)) or (easyPickCount > 9) or (not visor_easyPickCheckIdent("5bf66d", easyPickVisorId))
      if (easyPickTrigger):
        easyPickCount = 0
      end
      easyPickPoseIdx = easyPickCount
      easyPickPose = visor_getPose3d(easyPickVisorId, easyPickPoseIdx)
      visor_easyPickUpdate(easyPickVisorId, "counter", easyPickPoseIdx)
      # begin: URCap Program Node
      #   Source: SensoPart VISOR Robotic, 2.0.0, SensoPart Industriesensorik GmbH
      #   Type: Image Acquisition Pose
      $ 1648 "Image Acquisition Pose" "noBreak"
      if (easyPickTrigger):
        if (not easyPickAtImgAcq):
          movej(pose_trans(easyPickImgAcqPose,p[0.0000,0.0000,-0.0000,0.0000,0.0000,0.0000]),a=1.3963,v=1.0472,t=0.000000,r=0.000000)
          easyPickAtImgAcq = True
        end
        easyPickPose = easyPickFuncTrigger(easyPickVisorId, easyPickSetJob, easyPickJobName, easyPickArmMounted)
      end
      # end: URCap Program Node
      # begin: URCap Program Node
      #   Source: SensoPart VISOR Robotic, 2.0.0, SensoPart Industriesensorik GmbH
      #   Type: Object Detected
      $ 1649 "Object Detected" "noBreak"
      if (visor_partsFound(easyPickVisorId) > 0):
        $ 1650 "Open Gripper" "noBreak"
        # begin: URCap Program Node
        #   Source: Robotiq_Grippers, 1.8.4.4844, Robotiq Inc.
        #   Type: Gripper
        $ 1651 "Gripper Open (1)" "noBreak"
        if not(gripper_connected[0]):
          popup("Gripper 1 must be connected to run this program.", "No connection", False, True, True)
        end
        if not(rq_is_gripper_activated("1")):
          popup("Gripper 1 is not activated. Go to Installation tab > Gripper to activate it and run the program again.", "Not activated", False, True, True)
        end
        rq_set_pos_spd_for(0, 102, 77, "1")
        rq_wait_pos_spe_for_request(0, 102, 77, "1")
        rq_go_to("1")
        rq_wait("1")
        # end: URCap Program Node
        $ 1652 "MoveJ" "noBreak"
        $ 1653 "Waypoint_88" "noBreak"
        movej(get_inverse_kin(Waypoint_88_p, qnear=Waypoint_88_q), a=0.6981317007977318, v=0.5235987755982988)
        $ 1654 "Waypoint_87" "noBreak"
        movej(get_inverse_kin(Waypoint_87_p, qnear=Waypoint_87_q), a=0.6981317007977318, v=0.5235987755982988)
        $ 1655 "Waypoint_89" "noBreak"
        movej(get_inverse_kin(Waypoint_89_p, qnear=Waypoint_89_q), a=0.6981317007977318, v=0.5235987755982988)
        $ 1656 "MoveL" "noBreak"
        $ 1657 "Waypoint_90" "noBreak"
        movel(Waypoint_90_p, a=0.6, v=0.12)
        # begin: URCap Program Node
        #   Source: Robotiq_Grippers, 1.8.4.4844, Robotiq Inc.
        #   Type: Gripper
        $ 1658 "Gripper Close (1)" "noBreak"
        if not(gripper_connected[0]):
          popup("Gripper 1 must be connected to run this program.", "No connection", False, True, True)
        end
        if not(rq_is_gripper_activated("1")):
          popup("Gripper 1 is not activated. Go to Installation tab > Gripper to activate it and run the program again.", "Not activated", False, True, True)
        end
        rq_set_pos_spd_for(255, 0, 0, "1")
        rq_wait_pos_spe_for_request(255, 0, 0, "1")
        rq_go_to("1")
        rq_wait("1")
        # end: URCap Program Node
        $ 1659 "Waypoint_89" "noBreak"
        movel(Waypoint_89_p, a=0.6, v=0.12)
        $ 1663 "MoveJ" "noBreak"
        $ 1664 "Waypoint_94" "noBreak"
        movej(get_inverse_kin(Waypoint_94_p, qnear=Waypoint_94_q), a=1.3962634015954636, v=1.0471975511965976)
        $ 1665 "Waypoint_93" "noBreak"
        movej(get_inverse_kin(Waypoint_93_p, qnear=Waypoint_93_q), a=1.3962634015954636, v=1.0471975511965976)
        # begin: URCap Program Node
        #   Source: SensoPart VISOR Robotic, 2.0.0, SensoPart Industriesensorik GmbH
        #   Type: Approach Pose
        $ 1666 "Approach Pose" "noBreak"
        movej(pose_trans(easyPickPose,p[0.0000,0.0000,-0.0000,0.0000,0.0000,0.0000]),a=0.6981,v=0.5236,t=0.000000,r=0.000000)
        # end: URCap Program Node
        # begin: URCap Program Node
        #   Source: SensoPart VISOR Robotic, 2.0.0, SensoPart Industriesensorik GmbH
        #   Type: Target Pose
        $ 1667 "Target Pose" "noBreak"
        movel(pose_trans(easyPickPose,p[0.0000,0.0000,-0.0000,0.0000,0.0000,0.0000]),a=0.2000,v=0.1000,t=0.000000,r=0.000000)
        # end: URCap Program Node
        $ 1668 "Close Gripper" "noBreak"
        $ 1669 "current_pose≔get_actual_tcp_pose()" "noBreak"
        global current_pose= get_actual_tcp_pose ()
        $ 1670 "place_pose≔pose_trans(current_pose, offset)" "noBreak"
        global place_pose=pose_trans(current_pose, offset)
        $ 1671 "MoveJ" "noBreak"
        $ 1672 "place_pose" "noBreak"
        movej(place_pose, a=0.5235987755982988, v=0.3490658503988659)
        # begin: URCap Program Node
        #   Source: Robotiq_Grippers, 1.8.4.4844, Robotiq Inc.
        #   Type: Gripper
        $ 1673 "Gripper Open (1)" "noBreak"
        if not(gripper_connected[0]):
          popup("Gripper 1 must be connected to run this program.", "No connection", False, True, True)
        end
        if not(rq_is_gripper_activated("1")):
          popup("Gripper 1 is not activated. Go to Installation tab > Gripper to activate it and run the program again.", "Not activated", False, True, True)
        end
        rq_set_pos_spd_for(0, 0, 0, "1")
        rq_wait_pos_spe_for_request(0, 0, 0, "1")
        rq_go_to("1")
        rq_wait("1")
        # end: URCap Program Node
        # begin: URCap Program Node
        #   Source: SensoPart VISOR Robotic, 2.0.0, SensoPart Industriesensorik GmbH
        #   Type: Exit Pose
        $ 1674 "Exit Pose" "noBreak"
        movel(pose_trans(easyPickPose,p[0.0000,0.0000,-0.0000,0.0000,0.0000,0.0000]),a=0.2000,v=0.1200,t=0.000000,r=0.000000)
        # end: URCap Program Node
        easyPickObjTaken = True
      end
      # end: URCap Program Node
      # begin: URCap Program Node
      #   Source: SensoPart VISOR Robotic, 2.0.0, SensoPart Industriesensorik GmbH
      #   Type: No Object Detected
      $ 1675 "No Object Detected" "noBreak"
      if (visor_partsFound(easyPickVisorId) < 1):
        $ 1676 "Popup: No Container detected" "noBreak"
        popup("No Container detected", "Message", False, False, blocking=True)
        else:
      end
      # end: URCap Program Node
    end
    easyPickCount = easyPickCount + 1
    visor_easyPickUpdate(easyPickVisorId, "counter", easyPickCount)
    visor_easyPickSetIdent("5bf66d", easyPickVisorId)
    # end: URCap Program Node
  end
  visorFuncEasyPick_d789e5()
  # end: URCap Program Node
  $ 1677 "MoveJ"
  $ 1678 "Waypoint_95" "breakAfter"
  movej(get_inverse_kin(Waypoint_95_p, qnear=Waypoint_95_q), a=1.3962634015954636, v=1.0471975511965976)
  $ 1679 "Wait: 2.0"
  sleep(2.0)
  elif (7 == switch_1):
    $ 1680 "Case 7"
  elif (8 == switch_1):
    $ 1709 "Case 8"
  elif (11 == switch_1):
    $ 1742 "Case 11"
  elif (12 == switch_1):
    $ 1779 "Case 12"
  elif (15 == switch_1):
    $ 1830 "Case 15"
  elif (30 == switch_1):
    $ 1833 "Case 30"
  elif (31 == switch_1):
    $ 1866 "Case 31"
  elif (32 == switch_1):
    $ 1878 "Case 32"
  elif (33 == switch_1):
    $ 1919 "Case 33"
  elif (35 == switch_1):
    $ 1985 "Case 35"
    $ 1986 "Pick the powder container"
    # begin: URCap Program Node
    #   Source: SensoPart VISOR Robotic, 2.0.0, SensoPart Industriesensorik GmbH
    #   Type: VISOR Robotic App
    $ 1989 "VISOR Easy Pick"
    def visorFuncEasyPick_fbe43c():
      # begin: URCap Program Node
      #   Source: SensoPart VISOR Robotic, 2.0.0, SensoPart Industriesensorik GmbH
      #   Type: Easy Pick Setup
      $ 1990 "# 1 Setup" "noBreak"
      local easyPickVisorId = 1
      local easyPickArmMounted = True
      local easyPickSetJob = True
      local easyPickJobName = "Container"
      local easyPickAtImgAcq = False
      local easyPickImgAcqPose = cont_img_pose
      # end: URCap Program Node
      # begin: URCap Program Node
      #   Source: SensoPart VISOR Robotic, 2.0.0, SensoPart Industriesensorik GmbH
      #   Type: Process
      $ 1991 "Process" "noBreak"
      local easyPickObjTaken = False
      local easyPickTrigger = False
      local easyPickPoseIdx = 0
      local easyPickPose = p[0,0,0,0,0,0]
      def easyPickFuncTrigger(visorId, setJob, jobName, arm):
      if (setJob):
        visor_changeJob(visorId, jobName, 6000)
      end
      if (arm):
        visor_trigger(visorId, 6000, "arm")
      else:
        visor_trigger(visorId, 6000)
      end
      global easyPickParts=visor_partsFound(visorId)
      visor_easyPickUpdate(visorId, "parts", visor_partsFound(visorId))
      return visor_getPose3d(visorId, 0)
    end
    while (not easyPickObjTaken):
      easyPickTrigger = (easyPickCount >= visor_partsFound(easyPickVisorId)) or (easyPickCount > 9) or (not visor_easyPickCheckIdent("954e70", easyPickVisorId))
      if (easyPickTrigger):
        easyPickCount = 0
      end
      easyPickPoseIdx = easyPickCount
      easyPickPose = visor_getPose3d(easyPickVisorId, easyPickPoseIdx)
      visor_easyPickUpdate(easyPickVisorId, "counter", easyPickPoseIdx)
      # begin: URCap Program Node
      #   Source: SensoPart VISOR Robotic, 2.0.0, SensoPart Industriesensorik GmbH
      #   Type: Image Acquisition Pose
      $ 1992 "Image Acquisition Pose" "noBreak"
      if (easyPickTrigger):
        if (not easyPickAtImgAcq):
          movej(pose_trans(easyPickImgAcqPose,p[0.0000,0.0000,-0.0000,0.0000,0.0000,0.0000]),a=1.3963,v=1.0472,t=0.000000,r=0.000000)
          easyPickAtImgAcq = True
        end
        easyPickPose = easyPickFuncTrigger(easyPickVisorId, easyPickSetJob, easyPickJobName, easyPickArmMounted)
      end
      # end: URCap Program Node
      # begin: URCap Program Node
      #   Source: SensoPart VISOR Robotic, 2.0.0, SensoPart Industriesensorik GmbH
      #   Type: Object Detected
      $ 1993 "Object Detected" "noBreak"
      if (visor_partsFound(easyPickVisorId) > 0):
        $ 1994 "Open Gripper" "noBreak"
        # begin: URCap Program Node
        #   Source: Robotiq_Grippers, 1.8.4.4844, Robotiq Inc.
        #   Type: Gripper
        $ 1995 "Gripper Open (1)" "noBreak"
        if not(gripper_connected[0]):
          popup("Gripper 1 must be connected to run this program.", "No connection", False, True, True)
        end
        if not(rq_is_gripper_activated("1")):
          popup("Gripper 1 is not activated. Go to Installation tab > Gripper to activate it and run the program again.", "Not activated", False, True, True)
        end
        rq_set_pos_spd_for(0, 102, 77, "1")
        rq_wait_pos_spe_for_request(0, 102, 77, "1")
        rq_go_to("1")
        rq_wait("1")
        # end: URCap Program Node
        $ 1996 "MoveJ" "noBreak"
        $ 1997 "Waypoint_13" "noBreak"
        movej(get_inverse_kin(Waypoint_13_p, qnear=Waypoint_13_q), a=1.3962634015954636, v=1.0471975511965976)
        # begin: URCap Program Node
        #   Source: SensoPart VISOR Robotic, 2.0.0, SensoPart Industriesensorik GmbH
        #   Type: Approach Pose
        $ 1998 "Approach Pose" "noBreak"
        movej(pose_trans(easyPickPose,p[0.0000,0.0000,0.0500,0.0000,0.0000,0.0000]),a=1.3963,v=1.0472,t=0.000000,r=0.000000)
        # end: URCap Program Node
        # begin: URCap Program Node
        #   Source: SensoPart VISOR Robotic, 2.0.0, SensoPart Industriesensorik GmbH
        #   Type: Target Pose
        $ 1999 "Target Pose" "noBreak"
        movel(pose_trans(easyPickPose,p[0.0000,0.0000,-0.0000,0.0000,0.0000,0.0000]),a=0.5000,v=0.2500,t=0.000000,r=0.000000)
        # end: URCap Program Node
        $ 2000 "Close Gripper" "noBreak"
        # begin: URCap Program Node
        #   Source: Robotiq_Grippers, 1.8.4.4844, Robotiq Inc.
        #   Type: Gripper
        $ 2001 "Gripper Close (1)" "noBreak"
        if not(gripper_connected[0]):
          popup("Gripper 1 must be connected to run this program.", "No connection", False, True, True)
        end
        if not(rq_is_gripper_activated("1")):
          popup("Gripper 1 is not activated. Go to Installation tab > Gripper to activate it and run the program again.", "Not activated", False, True, True)
        end
        rq_set_pos_spd_for(255, 102, 77, "1")
        rq_wait_pos_spe_for_request(255, 102, 77, "1")
        rq_go_to("1")
        rq_wait("1")
        # end: URCap Program Node
        # begin: URCap Program Node
        #   Source: SensoPart VISOR Robotic, 2.0.0, SensoPart Industriesensorik GmbH
        #   Type: Exit Pose
        $ 2002 "Exit Pose" "noBreak"
        movel(pose_trans(easyPickPose,p[0.0000,0.0000,0.0500,0.0000,0.0000,0.0000]),a=0.5000,v=0.2500,t=0.000000,r=0.000000)
        # end: URCap Program Node
        easyPickObjTaken = True
      end
      # end: URCap Program Node
      # begin: URCap Program Node
      #   Source: SensoPart VISOR Robotic, 2.0.0, SensoPart Industriesensorik GmbH
      #   Type: No Object Detected
      $ 2003 "No Object Detected" "noBreak"
      if (visor_partsFound(easyPickVisorId) < 1):
        $ 2004 "Popup: No Container detected" "noBreak"
        popup("No Container detected", "Message", False, False, blocking=True)
        else:
      end
      # end: URCap Program Node
    end
    easyPickCount = easyPickCount + 1
    visor_easyPickUpdate(easyPickVisorId, "counter", easyPickCount)
    visor_easyPickSetIdent("954e70", easyPickVisorId)
    # end: URCap Program Node
  end
  visorFuncEasyPick_fbe43c()
  # end: URCap Program Node
  $ 2005 "MoveJ"
  $ 2007 "Waypoint_70" "breakAfter"
  movej(get_inverse_kin(Waypoint_70_p, qnear=Waypoint_70_q), a=0.6981317007977318, v=0.5235987755982988)
  $ 2008 "Waypoint_2" "breakAfter"
  movej(get_inverse_kin(Waypoint_2_p, qnear=Waypoint_2_q), a=0.8726646259971648, v=0.5235987755982988, r=0.05)
  $ 2009 "Waypoint_3" "breakAfter"
  movej(get_inverse_kin(Waypoint_3_p, qnear=Waypoint_3_q), a=0.6981317007977318, v=0.5235987755982988, r=0.05)
  $ 2010 "MoveL"
  $ 2011 "Waypoint_15" "breakAfter"
  movel(Waypoint_15_p, a=0.5, v=0.1, r=0.05)
  $ 2012 "Waypoint_14" "breakAfter"
  movel(Waypoint_14_p, a=0.3, v=0.1)
  $ 2013 "Waypoint_4" "breakAfter"
  movel(Waypoint_4_p, a=0.3, v=0.05)
  # begin: URCap Program Node
  #   Source: Robotiq_Grippers, 1.8.4.4844, Robotiq Inc.
  #   Type: Gripper
  $ 2014 "Gripper Open (1)"
  if not(gripper_connected[0]):
    popup("Gripper 1 must be connected to run this program.", "No connection", False, True, True)
  end
  if not(rq_is_gripper_activated("1")):
    popup("Gripper 1 is not activated. Go to Installation tab > Gripper to activate it and run the program again.", "Not activated", False, True, True)
  end
  rq_set_pos_spd_for(0, 102, 77, "1")
  rq_wait_pos_spe_for_request(0, 102, 77, "1")
  rq_go_to("1")
  rq_wait("1")
  # end: URCap Program Node
  $ 2015 "MoveL"
  $ 2016 "Waypoint_25" "breakAfter"
  movel(Waypoint_25_p, a=0.3, v=0.1)
  $ 2017 "Waypoint_15" "breakAfter"
  movel(Waypoint_15_p, a=0.5, v=0.1, r=0.05)
  $ 2018 "Home (Safe)"
  movej([-1.2302089344500047, -1.2969853503591224, -1.875639182904262, -1.539621866126728, 1.5731943360401213, -2.80099559440227], a=1.3962634015954636, v=1.0471975511965976)
  elif (36 == switch_1):
    $ 2048 "Case 36"
    $ 2052 "Decap"
    $ 2090 "MoveJ"
    $ 2091 "Waypoint_39" "breakAfter"
    movej(get_inverse_kin(Waypoint_39_p, qnear=Waypoint_39_q), a=1.3962634015954636, v=1.0471975511965976)
    $ 2092 "MoveL"
    $ 2093 "Waypoint_41" "breakAfter"
    movel(Waypoint_41_p, a=0.5, v=0.1)
    $ 2094 "Waypoint_40" "breakAfter"
    movel(Waypoint_40_p, a=0.3, v=0.05)
    # begin: URCap Program Node
    #   Source: Robotiq_Grippers, 1.8.4.4844, Robotiq Inc.
    #   Type: Gripper
    $ 2095 "Gripper Close (1)"
    if not(gripper_connected[0]):
      popup("Gripper 1 must be connected to run this program.", "No connection", False, True, True)
    end
    if not(rq_is_gripper_activated("1")):
      popup("Gripper 1 is not activated. Go to Installation tab > Gripper to activate it and run the program again.", "Not activated", False, True, True)
    end
    rq_set_pos_spd_for(255, 77, 51, "1")
    rq_wait_pos_spe_for_request(255, 77, 51, "1")
    rq_go_to("1")
    rq_wait("1")
    # end: URCap Program Node
    $ 2096 "Loop 2 times"
    Loop_2 = 0
    while (Loop_2 < 2):
      $ 2097 "MoveL"
      $ 2098 "Waypoint_42" "breakAfter"
      movel(Waypoint_42_p, a=1.2, v=0.5)
      $ 2099 "Waypoint_43" "breakAfter"
      movel(Waypoint_43_p, a=1.2, v=0.25)
      # begin: URCap Program Node
      #   Source: Robotiq_Grippers, 1.8.4.4844, Robotiq Inc.
      #   Type: Gripper
      $ 2100 "Gripper Move40mm (1)"
      if not(gripper_connected[0]):
        popup("Gripper 1 must be connected to run this program.", "No connection", False, True, True)
      end
      if not(rq_is_gripper_activated("1")):
        popup("Gripper 1 is not activated. Go to Installation tab > Gripper to activate it and run the program again.", "Not activated", False, True, True)
      end
      rq_set_pos_spd_for(63, 77, 51, "1")
      rq_wait_pos_spe_for_request(63, 77, 51, "1")
      rq_go_to("1")
      rq_wait("1")
      # end: URCap Program Node
      $ 2101 "MoveL"
      $ 2102 "Waypoint_44" "breakAfter"
      movel(Waypoint_44_p, a=1.2, v=0.5)
      $ 2103 "Waypoint_45" "breakAfter"
      movel(Waypoint_45_p, a=1.2, v=0.25)
      # begin: URCap Program Node
      #   Source: Robotiq_Grippers, 1.8.4.4844, Robotiq Inc.
      #   Type: Gripper
      $ 2104 "Gripper Move11mm (1)"
      if not(gripper_connected[0]):
        popup("Gripper 1 must be connected to run this program.", "No connection", False, True, True)
      end
      if not(rq_is_gripper_activated("1")):
        popup("Gripper 1 is not activated. Go to Installation tab > Gripper to activate it and run the program again.", "Not activated", False, True, True)
      end
      rq_set_pos_spd_for(200, 77, 51, "1")
      rq_wait_pos_spe_for_request(200, 77, 51, "1")
      rq_go_to("1")
      rq_wait("1")
      # end: URCap Program Node
      Loop_2 = Loop_2 + 1
    end
    $ 2105 "MoveL"
    $ 2106 "Waypoint_46" "breakAfter"
    movel(Waypoint_46_p, a=0.3, v=0.05)
    $ 2107 "Waypoint_47" "breakAfter"
    movel(Waypoint_47_p, a=0.5, v=0.1)
    $ 2108 "Waypoint_48" "breakAfter"
    movel(Waypoint_48_p, a=1.2, v=0.25)
    $ 2109 "Waypoint_49" "breakAfter"
    movel(Waypoint_49_p, a=1.2, v=0.25)
    # begin: URCap Program Node
    #   Source: Robotiq_Grippers, 1.8.4.4844, Robotiq Inc.
    #   Type: Gripper
    $ 2110 "Gripper Move35mm (1)"
    if not(gripper_connected[0]):
      popup("Gripper 1 must be connected to run this program.", "No connection", False, True, True)
    end
    if not(rq_is_gripper_activated("1")):
      popup("Gripper 1 is not activated. Go to Installation tab > Gripper to activate it and run the program again.", "Not activated", False, True, True)
    end
    rq_set_pos_spd_for(87, 77, 51, "1")
    rq_wait_pos_spe_for_request(87, 77, 51, "1")
    rq_go_to("1")
    rq_wait("1")
    # end: URCap Program Node
    $ 2111 "MoveL"
    $ 2112 "Waypoint_50" "breakAfter"
    movel(Waypoint_50_p, a=1.2, v=0.25)
    $ 2113 "Home (Safe)"
    movej([-1.2302089344500047, -1.2969853503591224, -1.875639182904262, -1.539621866126728, 1.5731943360401213, -2.80099559440227], a=1.3962634015954636, v=1.0471975511965976)
  elif (37 == switch_1):
    $ 2114 "Case 37"
  elif (38 == switch_1):
    $ 2248 "Case 38"
  elif (39 == switch_1):
    $ 2282 "Case 39"
  elif (40 == switch_1):
    $ 2334 "Case 40"
  end
  $ 2546 "'=========='"
  # '=========='
  $ 2547 "PostSettings"
  $ 2548 "'ADD ADDITIONAL CHECKS'"
  # 'ADD ADDITIONAL CHECKS'
  end
  $ 2 "BeforeStart"
  $ 3 "Scripts"
  $ 4 "Script: 001 SCRIPT Errors and Warnings Deifnes V0.2.script"

